  MoveL 4360 to (0, -14.4, 0.6) mm, rotated rx 0 ry 0 rz 180 deg; joints [18.174, -54.447, 108.401, -157.902, 56.008, 77.211]
  MoveL 4361 to (0, -15, 0.6) mm, rotated rx 0 ry 0 rz 180 deg; joints [18.174, -54.475, 108.395, -157.894, 55.977, 77.196]
  MoveL 4362 to (-200, -15, 0.6) mm, rotated rx 0 ry 0 rz 180 deg; joints [21.022, -63.449, 124.341, -156.258, 62.995, 78.705]
  MoveL 4363 to (-200, -15.6, 0.6) mm, rotated rx 0 ry 0 rz 180 deg; joints [21.022, -63.483, 124.335, -156.249, 62.958, 78.687]
  MoveL 4364 to (0, -15.6, 0.6) mm, rotated rx 0 ry 0 rz 180 deg; joints [18.174, -54.503, 108.39, -157.885, 55.945, 77.18]
  MoveL 4365 to (0, -16.2, 0.6) mm, rotated rx 0 ry 0 rz 180 deg; joints [18.174, -54.532, 108.384, -157.877, 55.914, 77.165]
  MoveL 4366 to (-200, -16.2, 0.6) mm, rotated rx 0 ry 0 rz 180 deg; joints [21.022, -63.518, 124.329, -156.241, 62.921, 78.669]
  MoveL 4367 to (-200, -16.8, 0.6) mm, rotated rx 0 ry 0 rz 180 deg; joints [21.022, -63.552, 124.323, -156.233, 62.883, 78.65]
  MoveL 4368 to (0, -16.8, 0.6) mm, rotated rx 0 ry 0 rz 180 deg; joints [18.174, -54.56, 108.378, -157.868, 55.882, 77.149]
  MoveL 4369 to (0, -17.4, 0.6) mm, rotated rx 0 ry 0 rz 180 deg; joints [18.174, -54.588, 108.373, -157.859, 55.851, 77.134]
  MoveL 4370 to (-200, -17.4, 0.6) mm, rotated rx 0 ry 0 rz 180 deg; joints [21.022, -63.586, 124.317, -156.224, 62.846, 78.632]
  MoveL 4371 to (-200, -18, 0.6) mm, rotated rx 0 ry 0 rz 180 deg; joints [21.022, -63.621, 124.311, -156.216, 62.809, 78.614]
  MoveL 4372 to (0, -18, 0.6) mm, rotated rx 0 ry 0 rz 180 deg; joints [18.174, -54.616, 108.367, -157.851, 55.819, 77.119]
  MoveL 4373 to (0, -18.6, 0.6) mm, rotated rx 0 ry 0 rz 180 deg; joints [18.174, -54.645, 108.361, -157.842, 55.788, 77.103]
  MoveL 4374 to (-200, -18.6, 0.6) mm, rotated rx 0 ry 0 rz 180 deg; joints [21.022, -63.655, 124.304, -156.208, 62.772, 78.595]
  MoveL 4375 to (-200, -19.2, 0.6) mm, rotated rx 0 ry 0 rz 180 deg; joints [21.022, -63.689, 124.298, -156.199, 62.735, 78.577]
  MoveL 4376 to (0, -19.2, 0.6) mm, rotated rx 0 ry 0 rz 180 deg; joints [18.174, -54.673, 108.355, -157.833, 55.756, 77.087]
  MoveL 4377 to (0, -19.8, 0.6) mm, rotated rx 0 ry 0 rz 180 deg; joints [18.174, -54.701, 108.349, -157.824, 55.725, 77.072]
  MoveL 4378 to (-200, -19.8, 0.6) mm, rotated rx 0 ry 0 rz 180 deg; joints [21.022, -63.724, 124.292, -156.191, 62.698, 78.558]
  MoveL 4379 to (-200, -20.4, 0.6) mm, rotated rx 0 ry 0 rz 180 deg; joints [21.022, -63.758, 124.285, -156.182, 62.661, 78.54]
  MoveL 4380 to (0, -20.4, 0.6) mm, rotated rx 0 ry 0 rz 180 deg; joints [18.174, -54.729, 108.344, -157.816, 55.693, 77.056]
  MoveL 4381 to (0, -21, 0.6) mm, rotated rx 0 ry 0 rz 180 deg; joints [18.174, -54.757, 108.338, -157.807, 55.662, 77.041]
  MoveL 4382 to (-200, -21, 0.6) mm, rotated rx 0 ry 0 rz 180 deg; joints [21.022, -63.792, 124.279, -156.174, 62.623, 78.521]
  MoveL 4383 to (-200, -21.6, 0.6) mm, rotated rx 0 ry 0 rz 180 deg; joints [21.022, -63.826, 124.272, -156.165, 62.586, 78.503]
  MoveL 4384 to (0, -21.6, 0.6) mm, rotated rx 0 ry 0 rz 180 deg; joints [18.174, -54.786, 108.332, -157.798, 55.63, 77.025]
  MoveL 4385 to (0, -22.2, 0.6) mm, rotated rx 0 ry 0 rz 180 deg; joints [18.174, -54.814, 108.326, -157.789, 55.599, 77.01]
  MoveL 4386 to (-200, -22.2, 0.6) mm, rotated rx 0 ry 0 rz 180 deg; joints [21.022, -63.86, 124.266, -156.157, 62.549, 78.484]
  MoveL 4387 to (-200, -22.8, 0.6) mm, rotated rx 0 ry 0 rz 180 deg; joints [21.022, -63.895, 124.26, -156.148, 62.512, 78.466]
  MoveL 4388 to (0, -22.8, 0.6) mm, rotated rx 0 ry 0 rz 180 deg; joints [18.174, -54.842, 108.32, -157.78, 55.567, 76.994]
  MoveL 4389 to (0, -23.4, 0.6) mm, rotated rx 0 ry 0 rz 180 deg; joints [18.174, -54.87, 108.314, -157.771, 55.535, 76.978]
  MoveL 4390 to (-200, -23.4, 0.6) mm, rotated rx 0 ry 0 rz 180 deg; joints [21.022, -63.929, 124.253, -156.14, 62.475, 78.447]
  MoveL 4391 to (-200, -24, 0.6) mm, rotated rx 0 ry 0 rz 180 deg; joints [21.022, -63.963, 124.246, -156.131, 62.438, 78.429]
  MoveL 4392 to (0, -24, 0.6) mm, rotated rx 0 ry 0 rz 180 deg; joints [18.174, -54.898, 108.308, -157.763, 55.504, 76.963]
  MoveL 4393 to (0, -24.6, 0.6) mm, rotated rx 0 ry 0 rz 180 deg; joints [18.174, -54.926, 108.302, -157.754, 55.472, 76.947]
  MoveL 4394 to (-200, -24.6, 0.6) mm, rotated rx 0 ry 0 rz 180 deg; joints [21.022, -63.997, 124.24, -156.122, 62.4, 78.41]
  MoveL 4395 to (-200, -25.2, 0.6) mm, rotated rx 0 ry 0 rz 180 deg; joints [21.022, -64.031, 124.233, -156.114, 62.363, 78.392]
  MoveL 4396 to (0, -25.2, 0.6) mm, rotated rx 0 ry 0 rz 180 deg; joints [18.174, -54.954, 108.296, -157.745, 55.441, 76.931]
  MoveL 4397 to (0, -25.8, 0.6) mm, rotated rx 0 ry 0 rz 180 deg; joints [18.174, -54.982, 108.289, -157.736, 55.409, 76.916]
  MoveL 4398 to (-200, -25.8, 0.6) mm, rotated rx 0 ry 0 rz 180 deg; joints [21.022, -64.065, 124.227, -156.105, 62.326, 78.373]
  MoveL 4399 to (-200, -26.4, 0.6) mm, rotated rx 0 ry 0 rz 180 deg; joints [21.022, -64.099, 124.22, -156.097, 62.289, 78.354]
  MoveL 4400 to (0, -26.4, 0.6) mm, rotated rx 0 ry 0 rz 180 deg; joints [18.174, -55.01, 108.283, -157.727, 55.377, 76.9]
  MoveL 4401 to (0, -27, 0.6) mm, rotated rx 0 ry 0 rz 180 deg; joints [18.174, -55.038, 108.277, -157.718, 55.346, 76.884]
  MoveL 4402 to (-200, -27, 0.6) mm, rotated rx 0 ry 0 rz 180 deg; joints [21.022, -64.133, 124.213, -156.088, 62.252, 78.336]
  MoveL 4403 to (-200, -27.6, 0.6) mm, rotated rx 0 ry 0 rz 180 deg; joints [21.022, -64.167, 124.206, -156.079, 62.214, 78.317]
  MoveL 4404 to (0, -27.6, 0.6) mm, rotated rx 0 ry 0 rz 180 deg; joints [18.174, -55.066, 108.271, -157.709, 55.314, 76.868]
  MoveL 4405 to (0, -28.2, 0.6) mm, rotated rx 0 ry 0 rz 180 deg; joints [18.174, -55.094, 108.265, -157.7, 55.282, 76.852]
  MoveL 4406 to (-200, -28.2, 0.6) mm, rotated rx 0 ry 0 rz 180 deg; joints [21.022, -64.201, 124.2, -156.07, 62.177, 78.298]
  MoveL 4407 to (-200, -28.8, 0.6) mm, rotated rx 0 ry 0 rz 180 deg; joints [21.022, -64.235, 124.193, -156.062, 62.14, 78.28]
  MoveL 4408 to (0, -28.8, 0.6) mm, rotated rx 0 ry 0 rz 180 deg; joints [18.174, -55.122, 108.258, -157.691, 55.251, 76.837]
  MoveL 4409 to (0, -29.4, 0.6) mm, rotated rx 0 ry 0 rz 180 deg; joints [18.174, -55.15, 108.252, -157.682, 55.219, 76.821]
  MoveL 4410 to (-200, -29.4, 0.6) mm, rotated rx 0 ry 0 rz 180 deg; joints [21.022, -64.269, 124.186, -156.053, 62.103, 78.261]
  MoveL 4411 to (-200, -30, 0.6) mm, rotated rx 0 ry 0 rz 180 deg; joints [21.022, -64.303, 124.179, -156.044, 62.065, 78.242]
  MoveL 4412 to (0, -30, 0.6) mm, rotated rx 0 ry 0 rz 180 deg; joints [18.174, -55.178, 108.246, -157.673, 55.187, 76.805]
  MoveL 4413 to (0, -30.6, 0.61) mm, rotated rx 2.39 ry 0 rz 180 deg; joints [18.094, -55.924, 108.131, -157.537, 54.374, 78.846]
  MoveL 4414 to (-200, -30.6, 0.61) mm, rotated rx 2.39 ry 0 rz 180 deg; joints [20.931, -65.205, 124.052, -155.918, 61.106, 80.201]
  MoveL 4415 to (-200, -31.2, 0.65) mm, rotated rx 4.78 ry 0 rz 180 deg; joints [20.813, -66.1, 123.923, -155.815, 60.147, 82.174]
  MoveL 4416 to (0, -31.2, 0.65) mm, rotated rx 4.78 ry 0 rz 180 deg; joints [17.989, -56.664, 108.016, -157.424, 53.559, 80.903]
  MoveL 4417 to (0, -31.8, 0.71) mm, rotated rx 7.16 ry 0 rz 180 deg; joints [17.861, -57.396, 107.901, -157.336, 52.745, 82.976]
  MoveL 4418 to (-200, -31.8, 0.71) mm, rotated rx 7.16 ry 0 rz 180 deg; joints [20.668, -66.984, 123.793, -155.736, 59.19, 84.161]
  MoveL 4419 to (-200, -32.39, 0.8) mm, rotated rx 9.55 ry 0 rz 180 deg; joints [20.495, -67.858, 123.663, -155.681, 58.234, 86.167]
  MoveL 4420 to (0, -32.39, 0.8) mm, rotated rx 9.55 ry 0 rz 180 deg; joints [17.708, -58.12, 107.785, -157.273, 51.933, 85.068]
  MoveL 4421 to (0, -32.98, 0.91) mm, rotated rx 11.94 ry 0 rz 180 deg; joints [17.531, -58.835, 107.67, -157.236, 51.122, 87.181]
  MoveL 4422 to (-200, -32.98, 0.91) mm, rotated rx 11.94 ry 0 rz 180 deg; joints [20.295, -68.721, 123.531, -155.653, 57.282, 88.193]
  MoveL 4423 to (-200, -33.56, 1.05) mm, rotated rx 14.32 ry 0 rz 180 deg; joints [20.068, -69.57, 123.4, -155.652, 56.333, 90.241]
  MoveL 4424 to (0, -33.56, 1.05) mm, rotated rx 14.32 ry 0 rz 180 deg; joints [17.331, -59.54, 107.555, -157.227, 50.315, 89.317]
  MoveL 4425 to (0, -34.14, 1.21) mm, rotated rx 16.71 ry 0 rz 180 deg; joints [17.107, -60.233, 107.441, -157.247, 49.513, 91.478]
  MoveL 4426 to (-200, -34.14, 1.21) mm, rotated rx 16.71 ry 0 rz 180 deg; joints [19.814, -70.405, 123.269, -155.68, 55.391, 92.314]
  MoveL 4427 to (-200, -34.71, 1.39) mm, rotated rx 19.1 ry 0 rz 180 deg; joints [19.533, -71.225, 123.138, -155.738, 54.454, 94.416]
  MoveL 4428 to (0, -34.71, 1.39) mm, rotated rx 19.1 ry 0 rz 180 deg; joints [16.859, -60.914, 107.328, -157.297, 48.715, 93.667]
  MoveL 4429 to (0, -35.27, 1.6) mm, rotated rx 21.49 ry 0 rz 180 deg; joints [16.589, -61.581, 107.218, -157.379, 47.925, 95.885]
  MoveL 4430 to (-200, -35.27, 1.6) mm, rotated rx 21.49 ry 0 rz 180 deg; joints [19.225, -72.028, 123.009, -155.827, 53.526, 96.546]
  MoveL 4431 to (-200, -35.83, 1.83) mm, rotated rx 23.87 ry 0 rz 180 deg; joints [18.892, -72.813, 122.882, -155.95, 52.606, 98.709]
  MoveL 4432 to (0, -35.83, 1.83) mm, rotated rx 23.87 ry 0 rz 180 deg; joints [16.295, -62.234, 107.109, -157.495, 47.142, 98.134]
  MoveL 4433 to (0, -36.37, 2.09) mm, rotated rx 26.26 ry 0 rz 180 deg; joints [15.979, -62.873, 107.003, -157.645, 46.368, 100.418]
  MoveL 4434 to (-200, -36.37, 2.09) mm, rotated rx 26.26 ry 0 rz 180 deg; joints [18.532, -73.58, 122.757, -156.107, 51.696, 100.907]
  MoveL 4435 to (-200, -36.9, 2.36) mm, rotated rx 28.65 ry 0 rz 180 deg; joints [18.147, -74.328, 122.635, -156.302, 50.798, 103.142]
  MoveL 4436 to (0, -36.9, 2.36) mm, rotated rx 28.65 ry 0 rz 180 deg; joints [15.641, -63.494, 106.9, -157.832, 45.604, 102.738]
  MoveL 4437 to (0, -37.42, 2.66) mm, rotated rx 31.03 ry 0 rz 180 deg; joints [15.281, -64.099, 106.8, -158.057, 44.853, 105.095]
  MoveL 4438 to (-200, -37.42, 2.66) mm, rotated rx 31.03 ry 0 rz 180 deg; joints [17.737, -75.054, 122.516, -156.535, 49.913, 105.418]
  MoveL 4439 to (-200, -37.93, 2.98) mm, rotated rx 33.42 ry 0 rz 180 deg; joints [17.301, -75.76, 122.401, -156.809, 49.042, 107.737]
  MoveL 4440 to (0, -37.93, 2.98) mm, rotated rx 33.42 ry 0 rz 180 deg; joints [14.9, -64.687, 106.705, -158.321, 44.114, 107.494]
  MoveL 4441 to (0, -38.42, 3.32) mm, rotated rx 35.81 ry 0 rz 180 deg; joints [14.498, -65.256, 106.613, -158.627, 43.39, 109.935]
  MoveL 4442 to (-200, -38.42, 3.32) mm, rotated rx 35.81 ry 0 rz 180 deg; joints [16.842, -76.442, 122.29, -157.125, 48.188, 110.1]
  MoveL 4443 to (-200, -38.91, 3.68) mm, rotated rx 38.2 ry 0 rz 180 deg; joints [16.358, -77.102, 122.185, -157.486, 47.352, 112.511]
  MoveL 4444 to (0, -38.91, 3.68) mm, rotated rx 38.2 ry 0 rz 180 deg; joints [14.076, -65.805, 106.527, -158.976, 42.682, 112.42]
  MoveL 4445 to (0, -39.37, 4.06) mm, rotated rx 40.59 ry 0 rz 180 deg; joints [13.634, -66.334, 106.446, -159.37, 41.992, 114.953]
  MoveL 4446 to (-200, -39.37, 4.06) mm, rotated rx 40.59 ry 0 rz 180 deg; joints [15.852, -77.737, 122.085, -157.893, 46.535, 114.973]
  MoveL 4447 to (-200, -39.82, 4.46) mm, rotated rx 42.97 ry 0 rz 180 deg; joints [15.322, -78.347, 121.991, -158.348, 45.739, 117.486]
  MoveL 4448 to (0, -39.82, 4.46) mm, rotated rx 42.97 ry 0 rz 180 deg; joints [13.173, -66.843, 106.37, -159.81, 41.321, 117.533]
  MoveL 4449 to (0, -40.25, 4.88) mm, rotated rx 45.36 ry 0 rz 180 deg; joints [12.693, -67.329, 106.301, -160.297, 40.672, 120.163]
  MoveL 4450 to (-200, -40.25, 4.88) mm, rotated rx 45.36 ry 0 rz 180 deg; joints [14.771, -78.931, 121.903, -158.853, 44.968, 120.054]
  MoveL 4451 to (-200, -40.66, 5.32) mm, rotated rx 47.75 ry 0 rz 180 deg; joints [14.199, -79.488, 121.823, -159.409, 44.222, 122.677]
  MoveL 4452 to (0, -40.66, 5.32) mm, rotated rx 47.75 ry 0 rz 180 deg; joints [12.196, -67.794, 106.238, -160.832, 40.045, 122.844]
  MoveL 4453 to (0, -41.05, 5.77) mm, rotated rx 50.13 ry 0 rz 180 deg; joints [11.681, -68.236, 106.182, -161.417, 39.444, 125.579]
  MoveL 4454 to (-200, -41.05, 5.77) mm, rotated rx 50.13 ry 0 rz 180 deg; joints [13.605, -80.018, 121.75, -160.019, 43.504, 125.36]
  MoveL 4455 to (-200, -41.43, 6.24) mm, rotated rx 52.52 ry 0 rz 180 deg; joints [12.993, -80.519, 121.685, -160.682, 42.817, 128.101]
  MoveL 4456 to (0, -41.43, 6.24) mm, rotated rx 52.52 ry 0 rz 180 deg; joints [11.15, -68.654, 106.134, -162.052, 38.869, 128.366]
  MoveL 4457 to (0, -41.78, 6.72) mm, rotated rx 54.91 ry 0 rz 180 deg; joints [10.604, -69.047, 106.093, -162.737, 38.324, 131.207]
  MoveL 4458 to (-200, -41.78, 6.72) mm, rotated rx 54.91 ry 0 rz 180 deg; joints [12.362, -80.992, 121.629, -161.4, 42.162, 130.901]
  MoveL 4459 to (-200, -42.12, 7.22) mm, rotated rx 57.3 ry 0 rz 180 deg; joints [11.713, -81.435, 121.582, -162.174, 41.541, 133.763]
  MoveL 4460 to (0, -42.12, 7.22) mm, rotated rx 57.3 ry 0 rz 180 deg; joints [10.043, -69.416, 106.061, -163.472, 37.809, 134.102]
  MoveL 4461 to (0, -42.43, 7.73) mm, rotated rx 59.68 ry 0 rz 180 deg; joints [9.469, -69.76, 106.037, -164.257, 37.327, 137.048]
  MoveL 4462 to (-200, -42.43, 7.73) mm, rotated rx 59.68 ry 0 rz 180 deg; joints [11.048, -81.848, 121.544, -163.002, 40.959, 136.684]
  MoveL 4463 to (-200, -42.72, 8.26) mm, rotated rx 62.07 ry 0 rz 180 deg; joints [10.368, -82.229, 121.516, -163.884, 40.416, 139.663]
  MoveL 4464 to (0, -42.72, 8.26) mm, rotated rx 62.07 ry 0 rz 180 deg; joints [8.883, -70.078, 106.021, -165.091, 36.88, 140.047]
  MoveL 4465 to (0, -42.99, 8.79) mm, rotated rx 64.46 ry 0 rz 180 deg; joints [8.284, -70.37, 106.015, -165.972, 36.47, 143.097]
  MoveL 4466 to (-200, -42.99, 8.79) mm, rotated rx 64.46 ry 0 rz 180 deg; joints [9.673, -82.58, 121.498, -164.82, 39.916, 142.702]
  MoveL 4467 to (-200, -43.24, 9.34) mm, rotated rx 66.84 ry 0 rz 180 deg; joints [8.965, -82.898, 121.49, -165.806, 39.461, 145.796]
  MoveL 4468 to (0, -43.24, 9.34) mm, rotated rx 66.84 ry 0 rz 180 deg; joints [7.675, -70.634, 106.017, -166.898, 36.099, 146.195]
  MoveL 4469 to (0, -43.46, 9.89) mm, rotated rx 69.23 ry 0 rz 180 deg; joints [7.057, -70.872, 106.029, -167.866, 35.769, 149.337]
  MoveL 4470 to (-200, -43.46, 9.89) mm, rotated rx 69.23 ry 0 rz 180 deg; joints [8.246, -83.184, 121.493, -166.841, 39.053, 148.942]
  MoveL 4471 to (-200, -43.66, 10.46) mm, rotated rx 71.62 ry 0 rz 180 deg; joints [7.517, -83.436, 121.507, -167.922, 38.695, 152.139]
  MoveL 4472 to (0, -43.66, 10.46) mm, rotated rx 71.62 ry 0 rz 180 deg; joints [6.431, -71.082, 106.051, -168.874, 35.481, 152.522]
  MoveL 4473 to (0, -43.84, 11.03) mm, rotated rx 74.01 ry 0 rz 180 deg; joints [5.797, -71.264, 106.082, -169.917, 35.237, 155.743]
  MoveL 4474 to (-200, -43.84, 11.03) mm, rotated rx 74.01 ry 0 rz 180 deg; joints [6.778, -83.656, 121.532, -169.044, 38.388, 155.379]
  MoveL 4475 to (-200, -44, 11.61) mm, rotated rx 76.39 ry 0 rz 180 deg; joints [6.032, -83.841, 121.568, -170.201, 38.135, 158.658]
  MoveL 4476 to (0, -44, 11.61) mm, rotated rx 76.39 ry 0 rz 180 deg; joints [5.158, -71.418, 106.123, -170.991, 35.039, 158.997]
  MoveL 4477 to (0, -44.12, 12.2) mm, rotated rx 78.78 ry 0 rz 180 deg; joints [4.514, -71.543, 106.173, -172.09, 34.887, 162.28]
  MoveL 4478 to (-200, -44.12, 12.2) mm, rotated rx 78.78 ry 0 rz 180 deg; joints [5.281, -83.992, 121.615, -171.391, 37.938, 161.973]
  MoveL 4479 to (-200, -44.23, 12.79) mm, rotated rx 81.17 ry 0 rz 180 deg; joints [4.525, -84.109, 121.674, -172.604, 37.797, 165.313]
  MoveL 4480 to (0, -44.23, 12.79) mm, rotated rx 81.17 ry 0 rz 180 deg; joints [3.867, -71.639, 106.234, -173.21, 34.783, 165.584]
  MoveL 4481 to (0, -44.31, 13.38) mm, rotated rx 83.56 ry 0 rz 180 deg; joints [3.218, -71.706, 106.304, -174.345, 34.728, 168.903]
  MoveL 4482 to (-200, -44.31, 13.38) mm, rotated rx 83.56 ry 0 rz 180 deg; joints [3.766, -84.191, 121.744, -173.836, 37.714, 168.673]
  MoveL 4483 to (-200, -44.36, 13.98) mm, rotated rx 85.94 ry 0 rz 180 deg; joints [3.006, -84.237, 121.825, -175.08, 37.69, 172.047]
  MoveL 4484 to (0, -44.36, 13.98) mm, rotated rx 85.94 ry 0 rz 180 deg; joints [2.568, -71.744, 106.384, -175.488, 34.722, 172.233]
  MoveL 4485 to (0, -44.39, 14.58) mm, rotated rx 88.33 ry 0 rz 180 deg; joints [1.919, -71.753, 106.473, -176.633, 34.766, 175.564]
  MoveL 4486 to (-200, -44.39, 14.58) mm, rotated rx 88.33 ry 0 rz 180 deg; joints [2.246, -84.249, 121.918, -176.328, 37.726, 175.425]
  MoveL 4487 to (-200, -44.4, 15.18) mm, rotated rx 90 ry 0 rz 180 deg; joints [1.707, -84.236, 121.989, -177.213, 37.786, 177.797]
  MoveL 4488 to (0, -44.4, 15.18) mm, rotated rx 90 ry 0 rz 180 deg; joints [1.459, -71.742, 106.541, -177.445, 34.826, 177.903]
  MoveL 4489 to (0, -44.4, 15.78) mm, rotated rx 90 ry 0 rz 180 deg; joints [1.433, -71.743, 106.542, -177.489, 34.825, 177.939]
  MoveL 4490 to (-200, -44.4, 15.78) mm, rotated rx 90 ry 0 rz 180 deg; joints [1.678, -84.237, 121.99, -177.261, 37.785, 177.834]
  MoveL 4491 to (-200, -44.4, 16.38) mm, rotated rx 90 ry 0 rz 180 deg; joints [1.649, -84.239, 121.992, -177.308, 37.784, 177.872]
  MoveL 4492 to (0, -44.4, 16.38) mm, rotated rx 90 ry 0 rz 180 deg; joints [1.408, -71.744, 106.544, -177.533, 34.825, 177.975]
  MoveL 4493 to (0, -44.4, 16.98) mm, rotated rx 90 ry 0 rz 180 deg; joints [1.383, -71.745, 106.545, -177.577, 34.824, 178.011]
  MoveL 4494 to (-200, -44.4, 16.98) mm, rotated rx 90 ry 0 rz 180 deg; joints [1.619, -84.24, 121.993, -177.356, 37.783, 177.91]
  MoveL 4495 to (-200, -44.4, 17.58) mm, rotated rx 90 ry 0 rz 180 deg; joints [1.59, -84.241, 121.994, -177.404, 37.782, 177.948]
  MoveL 4496 to (0, -44.4, 17.58) mm, rotated rx 90 ry 0 rz 180 deg; joints [1.358, -71.746, 106.546, -177.621, 34.824, 178.047]
  MoveL 4497 to (0, -44.4, 18.18) mm, rotated rx 90 ry 0 rz 180 deg; joints [1.333, -71.746, 106.547, -177.665, 34.823, 178.083]
  MoveL 4498 to (-200, -44.4, 18.18) mm, rotated rx 90 ry 0 rz 180 deg; joints [1.561, -84.242, 121.995, -177.452, 37.781, 177.986]
  MoveL 4499 to (-200, -44.4, 18.78) mm, rotated rx 90 ry 0 rz 180 deg; joints [1.531, -84.243, 121.996, -177.5, 37.78, 178.023]
  MoveL 4500 to (0, -44.4, 18.78) mm, rotated rx 90 ry 0 rz 180 deg; joints [1.308, -71.747, 106.548, -177.709, 34.823, 178.119]
  MoveL 4501 to (0, -44.4, 19.38) mm, rotated rx 90 ry 0 rz 180 deg; joints [1.283, -71.748, 106.549, -177.752, 34.822, 178.155]
  MoveL 4502 to (-200, -44.4, 19.38) mm, rotated rx 90 ry 0 rz 180 deg; joints [1.502, -84.244, 121.998, -177.548, 37.779, 178.061]
  MoveL 4503 to (-200, -44.4, 19.98) mm, rotated rx 90 ry 0 rz 180 deg; joints [1.473, -84.245, 121.999, -177.595, 37.778, 178.099]
  MoveL 4504 to (0, -44.4, 19.98) mm, rotated rx 90 ry 0 rz 180 deg; joints [1.258, -71.749, 106.551, -177.796, 34.822, 178.191]
  MoveL 4505 to (0, -44.4, 20.58) mm, rotated rx 90 ry 0 rz 180 deg; joints [1.233, -71.75, 106.552, -177.84, 34.821, 178.227]
  MoveL 4506 to (-200, -44.4, 20.58) mm, rotated rx 90 ry 0 rz 180 deg; joints [1.443, -84.246, 122, -177.643, 37.777, 178.137]
  MoveL 4507 to (-200, -44.4, 21.18) mm, rotated rx 90 ry 0 rz 180 deg; joints [1.414, -84.247, 122.001, -177.691, 37.777, 178.175]
  MoveL 4508 to (0, -44.4, 21.18) mm, rotated rx 90 ry 0 rz 180 deg; joints [1.208, -71.75, 106.553, -177.884, 34.821, 178.263]
  MoveL 4509 to (0, -44.4, 21.78) mm, rotated rx 90 ry 0 rz 180 deg; joints [1.183, -71.751, 106.554, -177.928, 34.82, 178.299]
  MoveL 4510 to (-200, -44.4, 21.78) mm, rotated rx 90 ry 0 rz 180 deg; joints [1.385, -84.248, 122.002, -177.739, 37.776, 178.212]
  MoveL 4511 to (-200, -44.4, 22.38) mm, rotated rx 90 ry 0 rz 180 deg; joints [1.356, -84.249, 122.003, -177.787, 37.775, 178.25]
  MoveL 4512 to (0, -44.4, 22.38) mm, rotated rx 90 ry 0 rz 180 deg; joints [1.158, -71.752, 106.555, -177.972, 34.82, 178.335]
  MoveL 4513 to (0, -44.4, 22.98) mm, rotated rx 90 ry 0 rz 180 deg; joints [1.133, -71.753, 106.556, -178.016, 34.819, 178.371]
  MoveL 4514 to (-200, -44.4, 22.98) mm, rotated rx 90 ry 0 rz 180 deg; joints [1.326, -84.25, 122.004, -177.835, 37.774, 178.288]
  MoveL 4515 to (-200, -44.4, 23.58) mm, rotated rx 90 ry 0 rz 180 deg; joints [1.297, -84.25, 122.005, -177.882, 37.773, 178.326]
  MoveL 4516 to (0, -44.4, 23.58) mm, rotated rx 90 ry 0 rz 180 deg; joints [1.108, -71.753, 106.557, -178.059, 34.819, 178.407]
  MoveL 4517 to (0, -44.4, 24.18) mm, rotated rx 90 ry 0 rz 180 deg; joints [1.083, -71.754, 106.558, -178.103, 34.818, 178.443]
  MoveL 4518 to (-200, -44.4, 24.18) mm, rotated rx 90 ry 0 rz 180 deg; joints [1.268, -84.251, 122.006, -177.93, 37.773, 178.364]
  MoveL 4519 to (-200, -44.4, 24.78) mm, rotated rx 90 ry 0 rz 180 deg; joints [1.238, -84.252, 122.007, -177.978, 37.772, 178.402]
  MoveL 4520 to (0, -44.4, 24.78) mm, rotated rx 90 ry 0 rz 180 deg; joints [1.058, -71.755, 106.559, -178.147, 34.818, 178.479]
  MoveL 4521 to (0, -44.4, 25.38) mm, rotated rx 90 ry 0 rz 180 deg; joints [1.033, -71.756, 106.56, -178.191, 34.817, 178.515]
  MoveL 4522 to (-200, -44.4, 25.38) mm, rotated rx 90 ry 0 rz 180 deg; joints [1.209, -84.253, 122.008, -178.026, 37.771, 178.439]
  MoveL 4523 to (-200, -44.4, 25.98) mm, rotated rx 90 ry 0 rz 180 deg; joints [1.18, -84.254, 122.009, -178.074, 37.77, 178.477]
  MoveL 4524 to (0, -44.4, 25.98) mm, rotated rx 90 ry 0 rz 180 deg; joints [1.008, -71.756, 106.56, -178.235, 34.817, 178.551]
  MoveL 4525 to (0, -44.4, 26.58) mm, rotated rx 90 ry 0 rz 180 deg; joints [0.983, -71.757, 106.561, -178.279, 34.817, 178.587]
  MoveL 4526 to (-200, -44.4, 26.58) mm, rotated rx 90 ry 0 rz 180 deg; joints [1.15, -84.255, 122.009, -178.122, 37.77, 178.515]
  MoveL 4527 to (-200, -44.4, 27.18) mm, rotated rx 90 ry 0 rz 180 deg; joints [1.121, -84.255, 122.01, -178.17, 37.769, 178.553]
  MoveL 4528 to (0, -44.4, 27.18) mm, rotated rx 90 ry 0 rz 180 deg; joints [0.958, -71.757, 106.562, -178.323, 34.816, 178.623]
  MoveL 4529 to (0, -44.4, 27.78) mm, rotated rx 90 ry 0 rz 180 deg; joints [0.933, -71.758, 106.563, -178.366, 34.816, 178.659]
  MoveL 4530 to (-200, -44.4, 27.78) mm, rotated rx 90 ry 0 rz 180 deg; joints [1.092, -84.256, 122.011, -178.217, 37.768, 178.591]
  MoveL 4531 to (-200, -44.4, 28.38) mm, rotated rx 90 ry 0 rz 180 deg; joints [1.062, -84.257, 122.012, -178.265, 37.768, 178.629]
  MoveL 4532 to (0, -44.4, 28.38) mm, rotated rx 90 ry 0 rz 180 deg; joints [0.907, -71.759, 106.564, -178.41, 34.815, 178.695]
  MoveL 4533 to (0, -44.4, 28.98) mm, rotated rx 90 ry 0 rz 180 deg; joints [0.882, -71.759, 106.565, -178.454, 34.815, 178.731]
  MoveL 4534 to (-200, -44.4, 28.98) mm, rotated rx 90 ry 0 rz 180 deg; joints [1.033, -84.258, 122.013, -178.313, 37.767, 178.666]
  MoveL 4535 to (-200, -44.4, 29.58) mm, rotated rx 90 ry 0 rz 180 deg; joints [1.004, -84.258, 122.014, -178.361, 37.767, 178.704]
  MoveL 4536 to (0, -44.4, 29.58) mm, rotated rx 90 ry 0 rz 180 deg; joints [0.857, -71.76, 106.565, -178.498, 34.815, 178.767]
  MoveL 4537 to (0, -44.4, 30.18) mm, rotated rx 90 ry 0 rz 180 deg; joints [0.832, -71.76, 106.566, -178.542, 34.814, 178.803]
  MoveL 4538 to (-200, -44.4, 30.18) mm, rotated rx 90 ry 0 rz 180 deg; joints [0.974, -84.259, 122.014, -178.409, 37.766, 178.742]
  MoveL 4539 to (-200, -44.4, 30.78) mm, rotated rx 90 ry 0 rz 180 deg; joints [0.945, -84.26, 122.015, -178.457, 37.766, 178.78]
  MoveL 4540 to (0, -44.4, 30.78) mm, rotated rx 90 ry 0 rz 180 deg; joints [0.807, -71.761, 106.567, -178.586, 34.814, 178.839]
  MoveL 4541 to (0, -44.4, 31.38) mm, rotated rx 90 ry 0 rz 180 deg; joints [0.782, -71.761, 106.567, -178.63, 34.814, 178.875]
  MoveL 4542 to (-200, -44.4, 31.38) mm, rotated rx 90 ry 0 rz 180 deg; joints [0.916, -84.26, 122.016, -178.505, 37.765, 178.818]
  MoveL 4543 to (-200, -44.4, 31.98) mm, rotated rx 90 ry 0 rz 180 deg; joints [0.886, -84.261, 122.016, -178.553, 37.764, 178.856]
  MoveL 4544 to (0, -44.4, 31.98) mm, rotated rx 90 ry 0 rz 180 deg; joints [0.757, -71.762, 106.568, -178.674, 34.813, 178.911]
  MoveL 4545 to (0, -44.4, 32.58) mm, rotated rx 90 ry 0 rz 180 deg; joints [0.732, -71.762, 106.569, -178.718, 34.813, 178.947]
  MoveL 4546 to (-200, -44.4, 32.58) mm, rotated rx 90 ry 0 rz 180 deg; joints [0.857, -84.261, 122.017, -178.6, 37.764, 178.894]
  MoveL 4547 to (-200, -44.4, 33.18) mm, rotated rx 90 ry 0 rz 180 deg; joints [0.828, -84.262, 122.018, -178.648, 37.763, 178.931]
  MoveL 4548 to (0, -44.4, 33.18) mm, rotated rx 90 ry 0 rz 180 deg; joints [0.707, -71.763, 106.569, -178.761, 34.813, 178.983]
  MoveL 4549 to (0, -44.4, 33.78) mm, rotated rx 90 ry 0 rz 180 deg; joints [0.682, -71.763, 106.57, -178.805, 34.813, 179.019]
  MoveL 4550 to (-200, -44.4, 33.78) mm, rotated rx 90 ry 0 rz 180 deg; joints [0.798, -84.262, 122.018, -178.696, 37.763, 178.969]
  MoveL 4551 to (-200, -44.4, 34.38) mm, rotated rx 90 ry 0 rz 180 deg; joints [0.769, -84.263, 122.019, -178.744, 37.763, 179.007]
  MoveL 4552 to (0, -44.4, 34.38) mm, rotated rx 90 ry 0 rz 180 deg; joints [0.657, -71.764, 106.571, -178.849, 34.812, 179.055]
  MoveL 4553 to (0, -44.4, 34.98) mm, rotated rx 90 ry 0 rz 180 deg; joints [0.632, -71.764, 106.571, -178.893, 34.812, 179.091]
  MoveL 4554 to (-200, -44.4, 34.98) mm, rotated rx 90 ry 0 rz 180 deg; joints [0.74, -84.263, 122.019, -178.792, 37.762, 179.045]
  MoveL 4555 to (-200, -44.4, 35.58) mm, rotated rx 90 ry 0 rz 180 deg; joints [0.71, -84.264, 122.02, -178.84, 37.762, 179.083]
  MoveL 4556 to (0, -44.4, 35.58) mm, rotated rx 90 ry 0 rz 180 deg; joints [0.607, -71.765, 106.572, -178.937, 34.812, 179.127]
  MoveL 4557 to (0, -44.4, 36.18) mm, rotated rx 90 ry 0 rz 180 deg; joints [0.582, -71.765, 106.572, -178.981, 34.812, 179.163]
  MoveL 4558 to (-200, -44.4, 36.18) mm, rotated rx 90 ry 0 rz 180 deg; joints [0.681, -84.264, 122.02, -178.888, 37.761, 179.121]
  MoveL 4559 to (-200, -44.4, 36.78) mm, rotated rx 90 ry 0 rz 180 deg; joints [0.652, -84.265, 122.021, -178.936, 37.761, 179.159]
  MoveL 4560 to (0, -44.4, 36.78) mm, rotated rx 90 ry 0 rz 180 deg; joints [0.557, -71.765, 106.573, -179.025, 34.811, 179.199]
  MoveL 4561 to (0, -44.4, 37.38) mm, rotated rx 90 ry 0 rz 180 deg; joints [0.532, -71.766, 106.573, -179.069, 34.811, 179.235]
  MoveL 4562 to (-200, -44.4, 37.38) mm, rotated rx 90 ry 0 rz 180 deg; joints [0.622, -84.265, 122.021, -178.984, 37.76, 179.196]
  MoveL 4563 to (-200, -44.4, 37.98) mm, rotated rx 90 ry 0 rz 180 deg; joints [0.593, -84.266, 122.022, -179.031, 37.76, 179.234]
  MoveL 4564 to (0, -44.4, 37.98) mm, rotated rx 90 ry 0 rz 180 deg; joints [0.507, -71.766, 106.574, -179.112, 34.811, 179.271]
  MoveL 4565 to (0, -44.4, 38.58) mm, rotated rx 90 ry 0 rz 180 deg; joints [0.482, -71.766, 106.574, -179.156, 34.811, 179.307]
  MoveL 4566 to (-200, -44.4, 38.58) mm, rotated rx 90 ry 0 rz 180 deg; joints [0.564, -84.266, 122.022, -179.079, 37.76, 179.272]
  MoveL 4567 to (-200, -44.4, 39.18) mm, rotated rx 90 ry 0 rz 180 deg; joints [0.534, -84.266, 122.023, -179.127, 37.759, 179.31]
  MoveL 4568 to (0, -44.4, 39.18) mm, rotated rx 90 ry 0 rz 180 deg; joints [0.457, -71.767, 106.574, -179.2, 34.81, 179.343]
  MoveL 4569 to (0, -44.4, 39.78) mm, rotated rx 90 ry 0 rz 180 deg; joints [0.431, -71.767, 106.575, -179.244, 34.81, 179.379]
  MoveL 4570 to (-200, -44.4, 39.78) mm, rotated rx 90 ry 0 rz 180 deg; joints [0.505, -84.267, 122.023, -179.175, 37.759, 179.348]
  MoveL 4571 to (-200, -44.4, 40.38) mm, rotated rx 90 ry 0 rz 180 deg; joints [0.476, -84.267, 122.024, -179.223, 37.759, 179.386]
  MoveL 4572 to (0, -44.4, 40.38) mm, rotated rx 90 ry 0 rz 180 deg; joints [0.406, -71.767, 106.575, -179.288, 34.81, 179.415]
  MoveL 4573 to (0, -44.4, 40.98) mm, rotated rx 90 ry 0 rz 180 deg; joints [0.381, -71.767, 106.576, -179.332, 34.81, 179.451]
  MoveL 4574 to (-200, -44.4, 40.98) mm, rotated rx 90 ry 0 rz 180 deg; joints [0.446, -84.267, 122.024, -179.271, 37.759, 179.424]
  MoveL 4575 to (-200, -44.4, 41.58) mm, rotated rx 90 ry 0 rz 180 deg; joints [0.417, -84.268, 122.024, -179.319, 37.758, 179.461]
  MoveL 4576 to (0, -44.4, 41.58) mm, rotated rx 90 ry 0 rz 180 deg; joints [0.356, -71.768, 106.576, -179.376, 34.81, 179.488]
  MoveL 4577 to (0, -44.4, 42.18) mm, rotated rx 90 ry 0 rz 180 deg; joints [0.331, -71.768, 106.576, -179.42, 34.81, 179.524]
  MoveL 4578 to (-200, -44.4, 42.18) mm, rotated rx 90 ry 0 rz 180 deg; joints [0.388, -84.268, 122.024, -179.367, 37.758, 179.499]
  MoveL 4579 to (-200, -44.4, 42.78) mm, rotated rx 90 ry 0 rz 180 deg; joints [0.358, -84.268, 122.025, -179.415, 37.758, 179.537]
  MoveL 4580 to (0, -44.4, 42.78) mm, rotated rx 90 ry 0 rz 180 deg; joints [0.306, -71.768, 106.576, -179.464, 34.81, 179.56]
  MoveL 4581 to (0, -44.4, 43.38) mm, rotated rx 90 ry 0 rz 180 deg; joints [0.281, -71.768, 106.577, -179.508, 34.809, 179.596]
  MoveL 4582 to (-200, -44.4, 43.38) mm, rotated rx 90 ry 0 rz 180 deg; joints [0.329, -84.269, 122.025, -179.463, 37.758, 179.575]
  MoveL 4583 to (-200, -44.4, 43.98) mm, rotated rx 90 ry 0 rz 180 deg; joints [0.3, -84.269, 122.025, -179.51, 37.758, 179.613]
  MoveL 4584 to (0, -44.4, 43.98) mm, rotated rx 90 ry 0 rz 180 deg; joints [0.256, -71.768, 106.577, -179.551, 34.809, 179.632]
  MoveL 4585 to (0, -44.4, 44.58) mm, rotated rx 90 ry 0 rz 180 deg; joints [0.231, -71.769, 106.577, -179.595, 34.809, 179.668]
  MoveL 4586 to (-200, -44.4, 44.58) mm, rotated rx 90 ry 0 rz 180 deg; joints [0.27, -84.269, 122.025, -179.558, 37.757, 179.651]
  MoveL 4587 to (-200, -44.4, 45.18) mm, rotated rx 90.72 ry 0 rz 180 deg; joints [0.022, -84.25, 122.049, -179.964, 37.799, -179.311]
  MoveL 4588 to (0, -44.4, 45.18) mm, rotated rx 90.72 ry 0 rz 180 deg; joints [0.019, -71.753, 106.599, -179.967, 34.846, -179.309]
  MoveL 4589 to (0, -44.38, 45.78) mm, rotated rx 93.11 ry 0 rz 180 deg; joints [-0.626, -71.682, 106.679, 178.909, 35.002, -176]
  MoveL 4590 to (-200, -44.38, 45.78) mm, rotated rx 93.11 ry 0 rz 180 deg; joints [-0.732, -84.166, 122.135, 178.81, 37.975, -175.956]
  MoveL 4591 to (-200, -44.33, 46.38) mm, rotated rx 95.49 ry 0 rz 180 deg; joints [-1.481, -84.045, 122.231, 177.605, 38.21, -172.625]
  MoveL 4592 to (0, -44.33, 46.38) mm, rotated rx 95.49 ry 0 rz 180 deg; joints [-1.265, -71.581, 106.767, 177.805, 35.206, -172.713]
  MoveL 4593 to (0, -44.26, 46.97) mm, rotated rx 97.88 ry 0 rz 180 deg; joints [-1.899, -71.451, 106.864, 176.725, 35.457, -169.452]
  MoveL 4594 to (-200, -44.26, 46.97) mm, rotated rx 97.88 ry 0 rz 180 deg; joints [-2.223, -83.89, 122.337, 176.428, 38.502, -169.323]
  MoveL 4595 to (-200, -44.17, 47.57) mm, rotated rx 100.27 ry 0 rz 180 deg; joints [-2.956, -83.699, 122.453, 175.284, 38.849, -166.056]
  MoveL 4596 to (0, -44.17, 47.57) mm, rotated rx 100.27 ry 0 rz 180 deg; joints [-2.526, -71.292, 106.97, 175.675, 35.755, -166.22]
  MoveL 4597 to (0, -44.05, 48.16) mm, rotated rx 102.66 ry 0 rz 180 deg; joints [-3.144, -71.104, 107.083, 174.659, 36.097, -163.025]
  MoveL 4598 to (-200, -44.05, 48.16) mm, rotated rx 102.66 ry 0 rz 180 deg; joints [-3.679, -83.474, 122.579, 174.18, 39.251, -162.832]
  MoveL 4599 to (-200, -43.91, 48.74) mm, rotated rx 105.04 ry 0 rz 180 deg; joints [-4.39, -83.213, 122.714, 173.119, 39.704, -159.653]
  MoveL 4600 to (0, -43.91, 48.74) mm, rotated rx 105.04 ry 0 rz 180 deg; joints [-3.752, -70.887, 107.204, 173.682, 36.483, -159.871]
  MoveL 4601 to (0, -43.74, 49.31) mm, rotated rx 107.43 ry 0 rz 180 deg; joints [-4.349, -70.642, 107.333, 172.745, 36.912, -156.758]
  MoveL 4602 to (-200, -43.74, 49.31) mm, rotated rx 107.43 ry 0 rz 180 deg; joints [-5.088, -82.918, 122.857, 172.104, 40.208, -156.524]
  MoveL 4603 to (-200, -43.55, 49.88) mm, rotated rx 109.82 ry 0 rz 180 deg; joints [-5.772, -82.589, 123.009, 171.139, 40.76, -153.448]
  MoveL 4604 to (0, -43.55, 49.88) mm, rotated rx 109.82 ry 0 rz 180 deg; joints [-4.935, -70.368, 107.468, 171.854, 37.379, -153.694]
  MoveL 4605 to (0, -43.33, 50.44) mm, rotated rx 112.2 ry 0 rz 180 deg; joints [-5.508, -70.067, 107.609, 171.008, 37.885, -150.677]
  MoveL 4606 to (-200, -43.33, 50.44) mm, rotated rx 112.2 ry 0 rz 180 deg; joints [-6.44, -82.226, 123.168, 170.227, 41.357, -150.429]
  MoveL 4607 to (-200, -43.09, 50.99) mm, rotated rx 114.59 ry 0 rz 180 deg; joints [-7.092, -81.829, 123.334, 169.367, 41.997, -147.465]
  MoveL 4608 to (0, -43.09, 50.99) mm, rotated rx 114.59 ry 0 rz 180 deg; joints [-6.066, -69.737, 107.756, 170.21, 38.428, -147.71]
  MoveL 4609 to (0, -42.83, 51.53) mm, rotated rx 116.98 ry 0 rz 180 deg; joints [-6.61, -69.381, 107.909, 169.462, 39.004, -144.795]
  MoveL 4610 to (-200, -42.83, 51.53) mm, rotated rx 116.98 ry 0 rz 180 deg; joints [-7.725, -81.4, 123.506, 168.563, 42.678, -144.561]
  MoveL 4611 to (-200, -42.55, 52.06) mm, rotated rx 119.37 ry 0 rz 180 deg; joints [-8.339, -80.938, 123.684, 167.814, 43.397, -141.716]
  MoveL 4612 to (0, -42.55, 52.06) mm, rotated rx 119.37 ry 0 rz 180 deg; joints [-7.137, -68.998, 108.066, 168.763, 39.612, -141.932]
  MoveL 4613 to (0, -42.24, 52.58) mm, rotated rx 121.75 ry 0 rz 180 deg; joints [-7.648, -68.588, 108.228, 168.114, 40.251, -139.12]
  MoveL 4614 to (-200, -42.24, 52.58) mm, rotated rx 121.75 ry 0 rz 180 deg; joints [-8.933, -80.444, 123.867, 167.119, 44.152, -138.928]
  MoveL 4615 to (-200, -41.92, 53.08) mm, rotated rx 124.14 ry 0 rz 180 deg; joints [-9.506, -79.918, 124.054, 166.479, 44.941, -136.199]
  MoveL 4616 to (0, -41.92, 53.08) mm, rotated rx 124.14 ry 0 rz 180 deg; joints [-8.141, -68.153, 108.393, 167.514, 40.917, -136.36]
  MoveL 4617 to (0, -41.57, 53.57) mm, rotated rx 126.53 ry 0 rz 180 deg; joints [-8.615, -67.692, 108.561, 166.963, 41.61, -133.65]
  MoveL 4618 to (-200, -41.57, 53.57) mm, rotated rx 126.53 ry 0 rz 180 deg; joints [-10.057, -79.362, 124.244, 165.892, 45.76, -133.526]
  MoveL 4619 to (-200, -41.2, 54.05) mm, rotated rx 128.92 ry 0 rz 180 deg; joints [-10.585, -78.775, 124.438, 165.357, 46.608, -130.908]
  MoveL 4620 to (0, -41.2, 54.05) mm, rotated rx 128.92 ry 0 rz 180 deg; joints [-9.07, -67.207, 108.731, 166.46, 42.326, -130.989]
  MoveL 4621 to (0, -40.82, 54.51) mm, rotated rx 131.3 ry 0 rz 180 deg; joints [-9.505, -66.699, 108.903, 166.005, 43.065, -128.377]
  MoveL 4622 to (-200, -40.82, 54.51) mm, rotated rx 131.3 ry 0 rz 180 deg; joints [-11.09, -78.16, 124.634, 164.873, 47.482, -128.343]
  MoveL 4623 to (-200, -40.41, 54.95) mm, rotated rx 133.69 ry 0 rz 180 deg; joints [-11.57, -77.515, 124.831, 164.438, 48.38, -125.83]
  MoveL 4624 to (0, -40.41, 54.95) mm, rotated rx 133.69 ry 0 rz 180 deg; joints [-9.919, -66.166, 109.076, 165.595, 43.823, -125.811]
  MoveL 4625 to (0, -39.99, 55.37) mm, rotated rx 136.08 ry 0 rz 180 deg; joints [-10.312, -65.612, 109.25, 165.229, 44.6, -123.29]
  MoveL 4626 to (-200, -39.99, 55.37) mm, rotated rx 136.08 ry 0 rz 180 deg; joints [-12.025, -76.843, 125.029, 164.05, 49.301, -123.366]
  MoveL 4627 to (-200, -39.55, 55.78) mm, rotated rx 138.47 ry 0 rz 180 deg; joints [-12.454, -76.144, 125.227, 163.708, 50.241, -120.947]
  MoveL 4628 to (0, -39.55, 55.78) mm, rotated rx 138.47 ry 0 rz 180 deg; joints [-10.684, -65.036, 109.424, 164.906, 45.394, -120.811]
  MoveL 4629 to (0, -39.09, 56.17) mm, rotated rx 140.85 ry 0 rz 180 deg; joints [-11.033, -64.438, 109.597, 164.625, 46.202, -118.373]
  MoveL 4630 to (-200, -39.09, 56.17) mm, rotated rx 140.85 ry 0 rz 180 deg; joints [-12.857, -75.419, 125.424, 163.409, 51.2, -118.573]
  MoveL 4631 to (-200, -38.62, 56.54) mm, rotated rx 143.24 ry 0 rz 180 deg; joints [-13.234, -74.669, 125.62, 163.153, 52.174, -116.241]
  MoveL 4632 to (0, -38.62, 56.54) mm, rotated rx 143.24 ry 0 rz 180 deg; joints [-11.359, -63.821, 109.769, 164.384, 47.024, -115.973]
  MoveL 4633 to (0, -38.13, 56.88) mm, rotated rx 145.63 ry 0 rz 180 deg; joints [-11.662, -63.185, 109.939, 164.18, 47.857, -113.608]
  MoveL 4634 to (-200, -38.13, 56.88) mm, rotated rx 145.63 ry 0 rz 180 deg; joints [-13.583, -73.895, 125.813, 162.936, 53.163, -113.945]
  MoveL 4635 to (-200, -37.63, 57.21) mm, rotated rx 148.01 ry 0 rz 180 deg; joints [-13.905, -73.099, 126.004, 162.757, 54.165, -111.687]
  MoveL 4636 to (0, -37.63, 57.21) mm, rotated rx 148.01 ry 0 rz 180 deg; joints [-11.941, -62.53, 110.107, 164.014, 48.7, -111.279]
  MoveL 4637 to (0, -37.11, 57.52) mm, rotated rx 150.4 ry 0 rz 180 deg; joints [-12.196, -61.858, 110.271, 163.882, 49.551, -108.981]
  MoveL 4638 to (-200, -37.11, 57.52) mm, rotated rx 150.4 ry 0 rz 180 deg; joints [-14.199, -72.28, 126.192, 162.615, 55.177, -109.462]
  MoveL 4639 to (-200, -36.59, 57.81) mm, rotated rx 152.79 ry 0 rz 180 deg; joints [-14.465, -71.441, 126.375, 162.507, 56.199, -107.266]
  MoveL 4640 to (0, -36.59, 57.81) mm, rotated rx 152.79 ry 0 rz 180 deg; joints [-12.427, -61.17, 110.433, 163.785, 50.409, -106.711]
  MoveL 4641 to (0, -36.05, 58.07) mm, rotated rx 155.18 ry 0 rz 180 deg; joints [-12.633, -60.466, 110.59, 163.719, 51.273, -104.47]
  MoveL 4642 to (-200, -36.05, 58.07) mm, rotated rx 155.18 ry 0 rz 180 deg; joints [-14.702, -70.583, 126.554, 162.432, 57.228, -105.1]
  MoveL 4643 to (-200, -35.5, 58.31) mm, rotated rx 157.56 ry 0 rz 180 deg; joints [-14.91, -69.707, 126.727, 162.389, 58.263, -102.958]
  MoveL 4644 to (0, -35.5, 58.31) mm, rotated rx 157.56 ry 0 rz 180 deg; joints [-12.814, -59.749, 110.743, 163.685, 52.141, -102.253]
  MoveL 4645 to (0, -34.94, 58.53) mm, rotated rx 159.95 ry 0 rz 180 deg; joints [-12.971, -59.018, 110.892, 163.68, 53.012, -100.058]
  MoveL 4646 to (-200, -34.94, 58.53) mm, rotated rx 159.95 ry 0 rz 180 deg; joints [-15.09, -68.814, 126.895, 162.377, 59.304, -100.838]
  MoveL 4647 to (-200, -34.37, 58.72) mm, rotated rx 162.34 ry 0 rz 180 deg; joints [-15.241, -67.906, 127.056, 162.393, 60.347, -98.739]
  MoveL 4648 to (0, -34.37, 58.72) mm, rotated rx 162.34 ry 0 rz 180 deg; joints [-13.102, -58.276, 111.035, 163.704, 53.885, -97.885]
  MoveL 4649 to (0, -33.79, 58.89) mm, rotated rx 164.72 ry 0 rz 180 deg; joints [-13.207, -57.523, 111.172, 163.755, 54.757, -95.73]
  MoveL 4650 to (-200, -33.79, 58.89) mm, rotated rx 164.72 ry 0 rz 180 deg; joints [-15.362, -66.984, 127.211, 162.437, 61.392, -96.657]
  MoveL 4651 to (-200, -33.21, 59.04) mm, rotated rx 167.11 ry 0 rz 180 deg; joints [-15.454, -66.049, 127.359, 162.507, 62.437, -94.59]
  MoveL 4652 to (0, -33.21, 59.04) mm, rotated rx 167.11 ry 0 rz 180 deg; joints [-13.288, -56.76, 111.304, 163.832, 55.629, -93.591]
  MoveL 4653 to (0, -32.62, 59.16) mm, rotated rx 169.5 ry 0 rz 180 deg; joints [-13.342, -55.99, 111.429, 163.934, 56.498, -91.468]
  MoveL 4654 to (-200, -32.62, 59.16) mm, rotated rx 169.5 ry 0 rz 180 deg; joints [-15.517, -65.104, 127.499, 162.604, 63.481, -92.537]
  MoveL 4655 to (-200, -32.03, 59.26) mm, rotated rx 171.89 ry 0 rz 180 deg; joints [-15.55, -64.15, 127.631, 162.725, 64.522, -90.494]
  MoveL 4656 to (0, -32.03, 59.26) mm, rotated rx 171.89 ry 0 rz 180 deg; joints [-13.371, -55.212, 111.548, 164.061, 57.364, -89.357]
  MoveL 4657 to (0, -31.44, 59.33) mm, rotated rx 174.28 ry 0 rz 180 deg; joints [-13.374, -54.429, 111.66, 164.212, 58.226, -87.257]
  MoveL 4658 to (-200, -31.44, 59.33) mm, rotated rx 174.28 ry 0 rz 180 deg; joints [-15.553, -63.188, 127.755, 162.871, 65.56, -88.458]
  MoveL 4659 to (-200, -30.84, 59.38) mm, rotated rx 176.66 ry 0 rz 180 deg; joints [-15.528, -62.221, 127.87, 163.04, 66.593, -86.43]
  MoveL 4660 to (0, -30.84, 59.38) mm, rotated rx 176.66 ry 0 rz 180 deg; joints [-13.352, -53.642, 111.765, 164.385, 59.082, -85.166]
  MoveL 4661 to (0, -30.24, 59.4) mm, rotated rx 179.05 ry 0 rz 180 deg; joints [-13.303, -52.852, 111.863, 164.58, 59.93, -83.083]
  MoveL 4662 to (-200, -30.24, 59.4) mm, rotated rx 179.05 ry 0 rz 180 deg; joints [-15.472, -61.249, 127.978, 163.232, 67.619, -84.406]
  MoveL 4663 to (-200, -29.64, 59.4) mm, rotated rx 180 ry 0 rz 180 deg; joints [-15.442, -60.838, 128.019, 163.317, 68.049, -83.608]
  MoveL 4664 to (0, -29.64, 59.4) mm, rotated rx 180 ry 0 rz 180 deg; joints [-13.277, -52.518, 111.902, 164.667, 60.286, -82.26]
  MoveL 4665 to (0, -29.04, 59.4) mm, rotated rx 180 ry 0 rz 180 deg; joints [-13.277, -52.486, 111.904, 164.672, 60.318, -82.271]
  MoveL 4666 to (-200, -29.04, 59.4) mm, rotated rx 180 ry 0 rz 180 deg; joints [-15.442, -60.799, 128.021, 163.322, 68.088, -83.62]
  MoveL 4667 to (-200, -28.44, 59.4) mm, rotated rx 180 ry 0 rz 180 deg; joints [-15.442, -60.761, 128.024, 163.326, 68.127, -83.633]
  MoveL 4668 to (0, -28.44, 59.4) mm, rotated rx 180 ry 0 rz 180 deg; joints [-13.277, -52.455, 111.906, 164.677, 60.35, -82.281]
  MoveL 4669 to (0, -27.84, 59.4) mm, rotated rx 180 ry 0 rz 180 deg; joints [-13.277, -52.424, 111.908, 164.682, 60.383, -82.291]
  MoveL 4670 to (-200, -27.84, 59.4) mm, rotated rx 180 ry 0 rz 180 deg; joints [-15.442, -60.722, 128.026, 163.331, 68.166, -83.646]
  MoveL 4671 to (-200, -27.24, 59.4) mm, rotated rx 180 ry 0 rz 180 deg; joints [-15.442, -60.684, 128.028, 163.336, 68.205, -83.658]
  MoveL 4672 to (0, -27.24, 59.4) mm, rotated rx 180 ry 0 rz 180 deg; joints [-13.277, -52.392, 111.91, 164.687, 60.415, -82.301]
  MoveL 4673 to (0, -26.64, 59.4) mm, rotated rx 180 ry 0 rz 180 deg; joints [-13.277, -52.361, 111.912, 164.692, 60.447, -82.311]
  MoveL 4674 to (-200, -26.64, 59.4) mm, rotated rx 180 ry 0 rz 180 deg; joints [-15.442, -60.645, 128.03, 163.34, 68.244, -83.671]
  MoveL 4675 to (-200, -26.04, 59.4) mm, rotated rx 180 ry 0 rz 180 deg; joints [-15.442, -60.607, 128.033, 163.345, 68.283, -83.683]
  MoveL 4676 to (0, -26.04, 59.4) mm, rotated rx 180 ry 0 rz 180 deg; joints [-13.277, -52.329, 111.914, 164.697, 60.479, -82.321]
  MoveL 4677 to (0, -25.44, 59.4) mm, rotated rx 180 ry 0 rz 180 deg; joints [-13.277, -52.298, 111.916, 164.702, 60.512, -82.332]
  MoveL 4678 to (-200, -25.44, 59.4) mm, rotated rx 180 ry 0 rz 180 deg; joints [-15.442, -60.568, 128.035, 163.35, 68.322, -83.696]
  MoveL 4679 to (-200, -24.84, 59.4) mm, rotated rx 180 ry 0 rz 180 deg; joints [-15.442, -60.529, 128.037, 163.354, 68.361, -83.709]
  MoveL 4680 to (0, -24.84, 59.4) mm, rotated rx 180 ry 0 rz 180 deg; joints [-13.277, -52.266, 111.918, 164.707, 60.544, -82.342]
  MoveL 4681 to (0, -24.24, 59.4) mm, rotated rx 180 ry 0 rz 180 deg; joints [-13.277, -52.235, 111.919, 164.712, 60.576, -82.352]
  MoveL 4682 to (-200, -24.24, 59.4) mm, rotated rx 180 ry 0 rz 180 deg; joints [-15.442, -60.491, 128.039, 163.359, 68.4, -83.721]
  MoveL 4683 to (-200, -23.64, 59.4) mm, rotated rx 180 ry 0 rz 180 deg; joints [-15.442, -60.452, 128.041, 163.364, 68.439, -83.734]
  MoveL 4684 to (0, -23.64, 59.4) mm, rotated rx 180 ry 0 rz 180 deg; joints [-13.277, -52.203, 111.921, 164.717, 60.608, -82.362]
  MoveL 4685 to (0, -23.04, 59.4) mm, rotated rx 180 ry 0 rz 180 deg; joints [-13.277, -52.172, 111.923, 164.722, 60.64, -82.372]
  MoveL 4686 to (-200, -23.04, 59.4) mm, rotated rx 180 ry 0 rz 180 deg; joints [-15.442, -60.414, 128.043, 163.368, 68.478, -83.746]
  MoveL 4687 to (-200, -22.44, 59.4) mm, rotated rx 180 ry 0 rz 180 deg; joints [-15.442, -60.375, 128.045, 163.373, 68.517, -83.759]
  MoveL 4688 to (0, -22.44, 59.4) mm, rotated rx 180 ry 0 rz 180 deg; joints [-13.277, -52.14, 111.925, 164.727, 60.672, -82.382]
  MoveL 4689 to (0, -21.84, 59.4) mm, rotated rx 180 ry 0 rz 180 deg; joints [-13.277, -52.109, 111.927, 164.732, 60.704, -82.392]
  MoveL 4690 to (-200, -21.84, 59.4) mm, rotated rx 180 ry 0 rz 180 deg; joints [-15.442, -60.336, 128.047, 163.377, 68.556, -83.771]
  MoveL 4691 to (-200, -21.24, 59.4) mm, rotated rx 180 ry 0 rz 180 deg; joints [-15.442, -60.297, 128.049, 163.382, 68.595, -83.784]
  MoveL 4692 to (0, -21.24, 59.4) mm, rotated rx 180 ry 0 rz 180 deg; joints [-13.277, -52.077, 111.928, 164.737, 60.737, -82.402]
  MoveL 4693 to (0, -20.64, 59.4) mm, rotated rx 180 ry 0 rz 180 deg; joints [-13.277, -52.046, 111.93, 164.742, 60.769, -82.412]
  MoveL 4694 to (-200, -20.64, 59.4) mm, rotated rx 180 ry 0 rz 180 deg; joints [-15.442, -60.259, 128.051, 163.387, 68.634, -83.796]
  MoveL 4695 to (-200, -20.04, 59.4) mm, rotated rx 180 ry 0 rz 180 deg; joints [-15.442, -60.22, 128.052, 163.391, 68.673, -83.809]
  MoveL 4696 to (0, -20.04, 59.4) mm, rotated rx 180 ry 0 rz 180 deg; joints [-13.277, -52.014, 111.932, 164.746, 60.801, -82.422]
  MoveL 4697 to (0, -19.44, 59.4) mm, rotated rx 180 ry 0 rz 180 deg; joints [-13.277, -51.982, 111.933, 164.751, 60.833, -82.432]
  MoveL 4698 to (-200, -19.44, 59.4) mm, rotated rx 180 ry 0 rz 180 deg; joints [-15.442, -60.181, 128.054, 163.396, 68.712, -83.821]
  MoveL 4699 to (-200, -18.84, 59.4) mm, rotated rx 180 ry 0 rz 180 deg; joints [-15.442, -60.142, 128.056, 163.4, 68.751, -83.833]
  MoveL 4700 to (0, -18.84, 59.4) mm, rotated rx 180 ry 0 rz 180 deg; joints [-13.277, -51.951, 111.935, 164.756, 60.865, -82.442]
  MoveL 4701 to (0, -18.24, 59.4) mm, rotated rx 180 ry 0 rz 180 deg; joints [-13.277, -51.919, 111.936, 164.761, 60.897, -82.452]
  MoveL 4702 to (-200, -18.24, 59.4) mm, rotated rx 180 ry 0 rz 180 deg; joints [-15.442, -60.104, 128.058, 163.405, 68.789, -83.846]
  MoveL 4703 to (-200, -17.64, 59.4) mm, rotated rx 180 ry 0 rz 180 deg; joints [-15.442, -60.065, 128.059, 163.409, 68.828, -83.858]
  MoveL 4704 to (0, -17.64, 59.4) mm, rotated rx 180 ry 0 rz 180 deg; joints [-13.277, -51.888, 111.938, 164.766, 60.929, -82.462]
  MoveL 4705 to (0, -17.04, 59.4) mm, rotated rx 180 ry 0 rz 180 deg; joints [-13.277, -51.856, 111.939, 164.771, 60.961, -82.472]
  MoveL 4706 to (-200, -17.04, 59.4) mm, rotated rx 180 ry 0 rz 180 deg; joints [-15.442, -60.026, 128.061, 163.414, 68.867, -83.871]
  MoveL 4707 to (-200, -16.44, 59.4) mm, rotated rx 180 ry 0 rz 180 deg; joints [-15.442, -59.987, 128.063, 163.418, 68.906, -83.883]
  MoveL 4708 to (0, -16.44, 59.4) mm, rotated rx 180 ry 0 rz 180 deg; joints [-13.277, -51.824, 111.941, 164.776, 60.993, -82.482]
  MoveL 4709 to (0, -15.84, 59.4) mm, rotated rx 180 ry 0 rz 180 deg; joints [-13.277, -51.792, 111.942, 164.78, 61.025, -82.492]
  MoveL 4710 to (-200, -15.84, 59.4) mm, rotated rx 180 ry 0 rz 180 deg; joints [-15.442, -59.948, 128.064, 163.422, 68.945, -83.895]
  MoveL 4711 to (-200, -15.24, 59.4) mm, rotated rx 180 ry 0 rz 180 deg; joints [-15.442, -59.909, 128.066, 163.427, 68.984, -83.908]
  MoveL 4712 to (0, -15.24, 59.4) mm, rotated rx 180 ry 0 rz 180 deg; joints [-13.277, -51.761, 111.944, 164.785, 61.057, -82.502]
  MoveL 4713 to (0, -14.64, 59.4) mm, rotated rx 180 ry 0 rz 180 deg; joints [-13.277, -51.729, 111.945, 164.79, 61.089, -82.512]
  MoveL 4714 to (-200, -14.64, 59.4) mm, rotated rx 180 ry 0 rz 180 deg; joints [-15.442, -59.87, 128.068, 163.431, 69.022, -83.92]
  MoveL 4715 to (-200, -14.04, 59.4) mm, rotated rx 180 ry 0 rz 180 deg; joints [-15.442, -59.831, 128.069, 163.436, 69.061, -83.933]
  MoveL 4716 to (0, -14.04, 59.4) mm, rotated rx 180 ry 0 rz 180 deg; joints [-13.277, -51.697, 111.947, 164.795, 61.121, -82.522]
  MoveL 4717 to (0, -13.44, 59.4) mm, rotated rx 180 ry 0 rz 180 deg; joints [-13.277, -51.665, 111.948, 164.8, 61.153, -82.532]
  MoveL 4718 to (-200, -13.44, 59.4) mm, rotated rx 180 ry 0 rz 180 deg; joints [-15.442, -59.792, 128.07, 163.44, 69.1, -83.945]
  MoveL 4719 to (-200, -12.84, 59.4) mm, rotated rx 180 ry 0 rz 180 deg; joints [-15.442, -59.753, 128.072, 163.445, 69.139, -83.957]
  MoveL 4720 to (0, -12.84, 59.4) mm, rotated rx 180 ry 0 rz 180 deg; joints [-13.277, -51.634, 111.949, 164.804, 61.185, -82.542]
  MoveL 4721 to (0, -12.24, 59.4) mm, rotated rx 180 ry 0 rz 180 deg; joints [-13.277, -51.602, 111.95, 164.809, 61.217, -82.552]
  MoveL 4722 to (-200, -12.24, 59.4) mm, rotated rx 180 ry 0 rz 180 deg; joints [-15.442, -59.714, 128.073, 163.449, 69.177, -83.97]
  MoveL 4723 to (-200, -11.64, 59.4) mm, rotated rx 180 ry 0 rz 180 deg; joints [-15.442, -59.675, 128.075, 163.453, 69.216, -83.982]
  MoveL 4724 to (0, -11.64, 59.4) mm, rotated rx 180 ry 0 rz 180 deg; joints [-13.277, -51.57, 111.952, 164.814, 61.249, -82.561]
  MoveL 4725 to (0, -11.04, 59.4) mm, rotated rx 180 ry 0 rz 180 deg; joints [-13.277, -51.538, 111.953, 164.819, 61.281, -82.571]
  MoveL 4726 to (-200, -11.04, 59.4) mm, rotated rx 180 ry 0 rz 180 deg; joints [-15.442, -59.636, 128.076, 163.458, 69.255, -83.994]
  MoveL 4727 to (-200, -10.44, 59.4) mm, rotated rx 180 ry 0 rz 180 deg; joints [-15.442, -59.597, 128.077, 163.462, 69.293, -84.006]
  MoveL 4728 to (0, -10.44, 59.4) mm, rotated rx 180 ry 0 rz 180 deg; joints [-13.277, -51.506, 111.954, 164.823, 61.312, -82.581]
  MoveL 4729 to (0, -9.84, 59.4) mm, rotated rx 180 ry 0 rz 180 deg; joints [-13.277, -51.474, 111.955, 164.828, 61.344, -82.591]
  MoveL 4730 to (-200, -9.84, 59.4) mm, rotated rx 180 ry 0 rz 180 deg; joints [-15.442, -59.558, 128.079, 163.466, 69.332, -84.019]
  MoveL 4731 to (-200, -9.24, 59.4) mm, rotated rx 180 ry 0 rz 180 deg; joints [-15.442, -59.519, 128.08, 163.471, 69.371, -84.031]
  MoveL 4732 to (0, -9.24, 59.4) mm, rotated rx 180 ry 0 rz 180 deg; joints [-13.277, -51.443, 111.956, 164.833, 61.376, -82.601]
  MoveL 4733 to (0, -8.64, 59.4) mm, rotated rx 180 ry 0 rz 180 deg; joints [-13.277, -51.411, 111.957, 164.838, 61.408, -82.611]
  MoveL 4734 to (-200, -8.64, 59.4) mm, rotated rx 180 ry 0 rz 180 deg; joints [-15.442, -59.48, 128.081, 163.475, 69.409, -84.043]
  MoveL 4735 to (-200, -8.04, 59.4) mm, rotated rx 180 ry 0 rz 180 deg; joints [-15.442, -59.441, 128.082, 163.479, 69.448, -84.055]
  MoveL 4736 to (0, -8.04, 59.4) mm, rotated rx 180 ry 0 rz 180 deg; joints [-13.277, -51.379, 111.959, 164.842, 61.44, -82.621]
  MoveL 4737 to (0, -7.44, 59.4) mm, rotated rx 180 ry 0 rz 180 deg; joints [-13.277, -51.347, 111.96, 164.847, 61.472, -82.63]
  MoveL 4738 to (-200, -7.44, 59.4) mm, rotated rx 180 ry 0 rz 180 deg; joints [-15.442, -59.402, 128.083, 163.484, 69.487, -84.068]
  MoveL 4739 to (-200, -6.84, 59.4) mm, rotated rx 180 ry 0 rz 180 deg; joints [-15.442, -59.363, 128.085, 163.488, 69.525, -84.08]
  MoveL 4740 to (0, -6.84, 59.4) mm, rotated rx 180 ry 0 rz 180 deg; joints [-13.277, -51.315, 111.961, 164.852, 61.503, -82.64]
  MoveL 4741 to (0, -6.24, 59.4) mm, rotated rx 180 ry 0 rz 180 deg; joints [-13.277, -51.283, 111.962, 164.856, 61.535, -82.65]
  MoveL 4742 to (-200, -6.24, 59.4) mm, rotated rx 180 ry 0 rz 180 deg; joints [-15.442, -59.323, 128.086, 163.492, 69.564, -84.092]
  MoveL 4743 to (-200, -5.64, 59.4) mm, rotated rx 180 ry 0 rz 180 deg; joints [-15.442, -59.284, 128.087, 163.496, 69.602, -84.104]
  MoveL 4744 to (0, -5.64, 59.4) mm, rotated rx 180 ry 0 rz 180 deg; joints [-13.277, -51.251, 111.962, 164.861, 61.567, -82.66]
  MoveL 4745 to (0, -5.04, 59.4) mm, rotated rx 180 ry 0 rz 180 deg; joints [-13.277, -51.219, 111.963, 164.866, 61.599, -82.669]
  MoveL 4746 to (-200, -5.04, 59.4) mm, rotated rx 180 ry 0 rz 180 deg; joints [-15.442, -59.245, 128.088, 163.501, 69.641, -84.116]
  MoveL 4747 to (-200, -4.44, 59.4) mm, rotated rx 180 ry 0 rz 180 deg; joints [-15.442, -59.206, 128.089, 163.505, 69.679, -84.129]
  MoveL 4748 to (0, -4.44, 59.4) mm, rotated rx 180 ry 0 rz 180 deg; joints [-13.277, -51.187, 111.964, 164.87, 61.63, -82.679]
  MoveL 4749 to (0, -3.84, 59.4) mm, rotated rx 180 ry 0 rz 180 deg; joints [-13.277, -51.155, 111.965, 164.875, 61.662, -82.689]
  MoveL 4750 to (-200, -3.84, 59.4) mm, rotated rx 180 ry 0 rz 180 deg; joints [-15.442, -59.167, 128.09, 163.509, 69.718, -84.141]
  MoveL 4751 to (-200, -3.24, 59.4) mm, rotated rx 180 ry 0 rz 180 deg; joints [-15.442, -59.127, 128.09, 163.513, 69.756, -84.153]
  MoveL 4752 to (0, -3.24, 59.4) mm, rotated rx 180 ry 0 rz 180 deg; joints [-13.277, -51.123, 111.966, 164.879, 61.694, -82.699]
  MoveL 4753 to (0, -2.64, 59.4) mm, rotated rx 180 ry 0 rz 180 deg; joints [-13.277, -51.091, 111.967, 164.884, 61.726, -82.708]
  MoveL 4754 to (-200, -2.64, 59.4) mm, rotated rx 180 ry 0 rz 180 deg; joints [-15.442, -59.088, 128.091, 163.517, 69.795, -84.165]
  MoveL 4755 to (-200, -2.04, 59.4) mm, rotated rx 180 ry 0 rz 180 deg; joints [-15.442, -59.049, 128.092, 163.522, 69.833, -84.177]
  MoveL 4756 to (0, -2.04, 59.4) mm, rotated rx 180 ry 0 rz 180 deg; joints [-13.277, -51.059, 111.967, 164.889, 61.757, -82.718]
  MoveL 4757 to (0, -1.44, 59.4) mm, rotated rx 180 ry 0 rz 180 deg; joints [-13.277, -51.027, 111.968, 164.893, 61.789, -82.728]
  MoveL 4758 to (-200, -1.44, 59.4) mm, rotated rx 180 ry 0 rz 180 deg; joints [-15.442, -59.01, 128.093, 163.526, 69.872, -84.189]
  MoveL 4759 to (-200, -0.84, 59.4) mm, rotated rx 180 ry 0 rz 180 deg; joints [-15.442, -58.97, 128.094, 163.53, 69.91, -84.201]
  MoveL 4760 to (0, -0.84, 59.4) mm, rotated rx 180 ry 0 rz 180 deg; joints [-13.277, -50.995, 111.969, 164.898, 61.821, -82.738]
  MoveL 4761 to (0, -0.24, 59.4) mm, rotated rx 180 ry 0 rz 180 deg; joints [-13.277, -50.962, 111.97, 164.902, 61.852, -82.747]
  MoveL 4762 to (-200, -0.24, 59.4) mm, rotated rx 180 ry 0 rz 180 deg; joints [-15.442, -58.931, 128.095, 163.534, 69.949, -84.214]
  MoveL 4763 to (-200, 0, 59.4) mm, rotated rx 180 ry 0 rz 180 deg; joints [-15.442, -58.915, 128.095, 163.536, 69.964, -84.218]
  MoveL 4764 to (0, 0, 59.4) mm, rotated rx 180 ry 0 rz 180 deg; joints [-13.277, -50.95, 111.97, 164.904, 61.865, -82.751]
  MoveL 4765 to (0, 0, 59.8) mm, rotated rx 180 ry 0 rz 180 deg; joints [-13.293, -50.946, 111.962, 164.886, 61.863, -82.741]
  MoveL 4766 to (-200, 0, 59.8) mm, rotated rx 180 ry 0 rz 180 deg; joints [-15.46, -58.911, 128.086, 163.516, 69.962, -84.21]
  MoveL 4767 to (-200, -0.6, 59.8) mm, rotated rx 180 ry 0 rz 180 deg; joints [-15.46, -58.95, 128.086, 163.512, 69.923, -84.198]
  MoveL 4768 to (0, -0.6, 59.8) mm, rotated rx 180 ry 0 rz 180 deg; joints [-13.293, -50.978, 111.961, 164.881, 61.831, -82.732]
  MoveL 4769 to (0, -1.2, 59.8) mm, rotated rx 180 ry 0 rz 180 deg; joints [-13.293, -51.01, 111.96, 164.877, 61.8, -82.722]
  MoveL 4770 to (-200, -1.2, 59.8) mm, rotated rx 180 ry 0 rz 180 deg; joints [-15.46, -58.99, 128.085, 163.508, 69.885, -84.186]
  MoveL 4771 to (-200, -1.8, 59.8) mm, rotated rx 180 ry 0 rz 180 deg; joints [-15.46, -59.029, 128.084, 163.504, 69.847, -84.174]
  MoveL 4772 to (0, -1.8, 59.8) mm, rotated rx 180 ry 0 rz 180 deg; joints [-13.293, -51.042, 111.96, 164.872, 61.768, -82.712]
  MoveL 4773 to (0, -2.4, 59.8) mm, rotated rx 180 ry 0 rz 180 deg; joints [-13.293, -51.074, 111.959, 164.868, 61.736, -82.703]
  MoveL 4774 to (-200, -2.4, 59.8) mm, rotated rx 180 ry 0 rz 180 deg; joints [-15.46, -59.068, 128.083, 163.499, 69.808, -84.162]
  MoveL 4775 to (-200, -3, 59.8) mm, rotated rx 180 ry 0 rz 180 deg; joints [-15.46, -59.108, 128.082, 163.495, 69.77, -84.15]
  MoveL 4776 to (0, -3, 59.8) mm, rotated rx 180 ry 0 rz 180 deg; joints [-13.293, -51.106, 111.958, 164.863, 61.705, -82.693]
  MoveL 4777 to (0, -3.6, 59.8) mm, rotated rx 180 ry 0 rz 180 deg; joints [-13.293, -51.138, 111.957, 164.858, 61.673, -82.683]
  MoveL 4778 to (-200, -3.6, 59.8) mm, rotated rx 180 ry 0 rz 180 deg; joints [-15.46, -59.147, 128.081, 163.491, 69.731, -84.138]
  MoveL 4779 to (-200, -4.2, 59.8) mm, rotated rx 180 ry 0 rz 180 deg; joints [-15.46, -59.186, 128.081, 163.487, 69.693, -84.126]
  MoveL 4780 to (0, -4.2, 59.8) mm, rotated rx 180 ry 0 rz 180 deg; joints [-13.293, -51.17, 111.957, 164.854, 61.641, -82.673]
  MoveL 4781 to (0, -4.8, 59.8) mm, rotated rx 180 ry 0 rz 180 deg; joints [-13.293, -51.202, 111.956, 164.849, 61.61, -82.664]
  MoveL 4782 to (-200, -4.8, 59.8) mm, rotated rx 180 ry 0 rz 180 deg; joints [-15.46, -59.225, 128.08, 163.483, 69.654, -84.113]
  MoveL 4783 to (-200, -5.4, 59.8) mm, rotated rx 180 ry 0 rz 180 deg; joints [-15.46, -59.264, 128.079, 163.478, 69.616, -84.101]
  MoveL 4784 to (0, -5.4, 59.8) mm, rotated rx 180 ry 0 rz 180 deg; joints [-13.293, -51.234, 111.955, 164.844, 61.578, -82.654]
  MoveL 4785 to (0, -6, 59.8) mm, rotated rx 180 ry 0 rz 180 deg; joints [-13.293, -51.266, 111.954, 164.84, 61.546, -82.644]
  MoveL 4786 to (-200, -6, 59.8) mm, rotated rx 180 ry 0 rz 180 deg; joints [-15.46, -59.304, 128.078, 163.474, 69.577, -84.089]
  MoveL 4787 to (-200, -6.6, 59.8) mm, rotated rx 180 ry 0 rz 180 deg; joints [-15.46, -59.343, 128.076, 163.47, 69.538, -84.077]
  MoveL 4788 to (0, -6.6, 59.8) mm, rotated rx 180 ry 0 rz 180 deg; joints [-13.293, -51.298, 111.953, 164.835, 61.514, -82.634]
  MoveL 4789 to (0, -7.2, 59.8) mm, rotated rx 180 ry 0 rz 180 deg; joints [-13.293, -51.33, 111.952, 164.83, 61.482, -82.624]
  MoveL 4790 to (-200, -7.2, 59.8) mm, rotated rx 180 ry 0 rz 180 deg; joints [-15.46, -59.382, 128.075, 163.466, 69.5, -84.064]
  MoveL 4791 to (-200, -7.8, 59.8) mm, rotated rx 180 ry 0 rz 180 deg; joints [-15.46, -59.421, 128.074, 163.461, 69.461, -84.052]
  MoveL 4792 to (0, -7.8, 59.8) mm, rotated rx 180 ry 0 rz 180 deg; joints [-13.293, -51.362, 111.951, 164.826, 61.451, -82.615]
  MoveL 4793 to (0, -8.4, 59.8) mm, rotated rx 180 ry 0 rz 180 deg; joints [-13.293, -51.394, 111.95, 164.821, 61.419, -82.605]
  MoveL 4794 to (-200, -8.4, 59.8) mm, rotated rx 180 ry 0 rz 180 deg; joints [-15.46, -59.46, 128.073, 163.457, 69.423, -84.04]
  MoveL 4795 to (-200, -9, 59.8) mm, rotated rx 180 ry 0 rz 180 deg; joints [-15.46, -59.499, 128.072, 163.453, 69.384, -84.028]
  MoveL 4796 to (0, -9, 59.8) mm, rotated rx 180 ry 0 rz 180 deg; joints [-13.293, -51.426, 111.949, 164.816, 61.387, -82.595]
  MoveL 4797 to (0, -9.6, 59.8) mm, rotated rx 180 ry 0 rz 180 deg; joints [-13.293, -51.458, 111.948, 164.812, 61.355, -82.585]
  MoveL 4798 to (-200, -9.6, 59.8) mm, rotated rx 180 ry 0 rz 180 deg; joints [-15.46, -59.538, 128.071, 163.448, 69.345, -84.015]
  MoveL 4799 to (-200, -10.2, 59.8) mm, rotated rx 180 ry 0 rz 180 deg; joints [-15.46, -59.577, 128.069, 163.444, 69.307, -84.003]
  MoveL 4800 to (0, -10.2, 59.8) mm, rotated rx 180 ry 0 rz 180 deg; joints [-13.293, -51.49, 111.946, 164.807, 61.323, -82.575]
  MoveL 4801 to (0, -10.8, 59.8) mm, rotated rx 180 ry 0 rz 180 deg; joints [-13.293, -51.521, 111.945, 164.802, 61.291, -82.565]
  MoveL 4802 to (-200, -10.8, 59.8) mm, rotated rx 180 ry 0 rz 180 deg; joints [-15.46, -59.617, 128.068, 163.44, 69.268, -83.991]
  MoveL 4803 to (-200, -11.4, 59.8) mm, rotated rx 180 ry 0 rz 180 deg; joints [-15.46, -59.656, 128.067, 163.435, 69.229, -83.979]
  MoveL 4804 to (0, -11.4, 59.8) mm, rotated rx 180 ry 0 rz 180 deg; joints [-13.293, -51.553, 111.944, 164.797, 61.26, -82.556]
  MoveL 4805 to (0, -12, 59.8) mm, rotated rx 180 ry 0 rz 180 deg; joints [-13.293, -51.585, 111.943, 164.793, 61.228, -82.546]
  MoveL 4806 to (-200, -12, 59.8) mm, rotated rx 180 ry 0 rz 180 deg; joints [-15.46, -59.695, 128.065, 163.431, 69.191, -83.966]
  MoveL 4807 to (-200, -12.6, 59.8) mm, rotated rx 180 ry 0 rz 180 deg; joints [-15.46, -59.734, 128.064, 163.427, 69.152, -83.954]
  MoveL 4808 to (0, -12.6, 59.8) mm, rotated rx 180 ry 0 rz 180 deg; joints [-13.293, -51.617, 111.942, 164.788, 61.196, -82.536]
  MoveL 4809 to (0, -13.2, 59.8) mm, rotated rx 180 ry 0 rz 180 deg; joints [-13.293, -51.649, 111.94, 164.783, 61.164, -82.526]
  MoveL 4810 to (-200, -13.2, 59.8) mm, rotated rx 180 ry 0 rz 180 deg; joints [-15.46, -59.773, 128.063, 163.422, 69.113, -83.942]
  MoveL 4811 to (-200, -13.8, 59.8) mm, rotated rx 180 ry 0 rz 180 deg; joints [-15.46, -59.811, 128.061, 163.418, 69.074, -83.929]
  MoveL 4812 to (0, -13.8, 59.8) mm, rotated rx 180 ry 0 rz 180 deg; joints [-13.293, -51.68, 111.939, 164.778, 61.132, -82.516]
  MoveL 4813 to (0, -14.4, 59.8) mm, rotated rx 180 ry 0 rz 180 deg; joints [-13.293, -51.712, 111.938, 164.773, 61.1, -82.506]
  MoveL 4814 to (-200, -14.4, 59.8) mm, rotated rx 180 ry 0 rz 180 deg; joints [-15.46, -59.85, 128.06, 163.413, 69.036, -83.917]
  MoveL 4815 to (-200, -15, 59.8) mm, rotated rx 180 ry 0 rz 180 deg; joints [-15.46, -59.889, 128.058, 163.409, 68.997, -83.905]
  MoveL 4816 to (0, -15, 59.8) mm, rotated rx 180 ry 0 rz 180 deg; joints [-13.293, -51.744, 111.936, 164.769, 61.068, -82.496]
  MoveL 4817 to (0, -15.6, 59.8) mm, rotated rx 180 ry 0 rz 180 deg; joints [-13.293, -51.776, 111.935, 164.764, 61.036, -82.486]
  MoveL 4818 to (-200, -15.6, 59.8) mm, rotated rx 180 ry 0 rz 180 deg; joints [-15.46, -59.928, 128.057, 163.404, 68.958, -83.892]
  MoveL 4819 to (-200, -16.2, 59.8) mm, rotated rx 180 ry 0 rz 180 deg; joints [-15.46, -59.967, 128.055, 163.4, 68.919, -83.88]
  MoveL 4820 to (0, -16.2, 59.8) mm, rotated rx 180 ry 0 rz 180 deg; joints [-13.293, -51.807, 111.933, 164.759, 61.004, -82.476]
  MoveL 4821 to (0, -16.8, 59.8) mm, rotated rx 180 ry 0 rz 180 deg; joints [-13.293, -51.839, 111.932, 164.754, 60.972, -82.466]
  MoveL 4822 to (-200, -16.8, 59.8) mm, rotated rx 180 ry 0 rz 180 deg; joints [-15.46, -60.006, 128.053, 163.396, 68.881, -83.867]
  MoveL 4823 to (-200, -17.4, 59.8) mm, rotated rx 180 ry 0 rz 180 deg; joints [-15.46, -60.045, 128.052, 163.391, 68.842, -83.855]
  MoveL 4824 to (0, -17.4, 59.8) mm, rotated rx 180 ry 0 rz 180 deg; joints [-13.293, -51.871, 111.931, 164.749, 60.94, -82.456]
  MoveL 4825 to (0, -18, 59.8) mm, rotated rx 180 ry 0 rz 180 deg; joints [-13.293, -51.902, 111.929, 164.744, 60.908, -82.446]
  MoveL 4826 to (-200, -18, 59.8) mm, rotated rx 180 ry 0 rz 180 deg; joints [-15.46, -60.084, 128.05, 163.387, 68.803, -83.843]
  MoveL 4827 to (-200, -18.6, 59.8) mm, rotated rx 180 ry 0 rz 180 deg; joints [-15.46, -60.123, 128.048, 163.382, 68.764, -83.83]
  MoveL 4828 to (0, -18.6, 59.8) mm, rotated rx 180 ry 0 rz 180 deg; joints [-13.293, -51.934, 111.927, 164.74, 60.876, -82.436]
  MoveL 4829 to (0, -19.2, 59.8) mm, rotated rx 180 ry 0 rz 180 deg; joints [-13.293, -51.966, 111.926, 164.735, 60.844, -82.426]
  MoveL 4830 to (-200, -19.2, 59.8) mm, rotated rx 180 ry 0 rz 180 deg; joints [-15.46, -60.161, 128.047, 163.378, 68.725, -83.818]
  MoveL 4831 to (-200, -19.8, 59.8) mm, rotated rx 180 ry 0 rz 180 deg; joints [-15.46, -60.2, 128.045, 163.373, 68.686, -83.805]
  MoveL 4832 to (0, -19.8, 59.8) mm, rotated rx 180 ry 0 rz 180 deg; joints [-13.293, -51.997, 111.924, 164.73, 60.812, -82.416]
  MoveL 4833 to (0, -20.4, 59.8) mm, rotated rx 180 ry 0 rz 180 deg; joints [-13.293, -52.029, 111.923, 164.725, 60.78, -82.406]
  MoveL 4834 to (-200, -20.4, 59.8) mm, rotated rx 180 ry 0 rz 180 deg; joints [-15.46, -60.239, 128.043, 163.368, 68.647, -83.793]
  MoveL 4835 to (-200, -21, 59.8) mm, rotated rx 180 ry 0 rz 180 deg; joints [-15.46, -60.278, 128.041, 163.364, 68.609, -83.78]
  MoveL 4836 to (0, -21, 59.8) mm, rotated rx 180 ry 0 rz 180 deg; joints [-13.293, -52.061, 111.921, 164.72, 60.748, -82.396]
  MoveL 4837 to (0, -21.6, 59.8) mm, rotated rx 180 ry 0 rz 180 deg; joints [-13.293, -52.092, 111.919, 164.715, 60.716, -82.386]
  MoveL 4838 to (-200, -21.6, 59.8) mm, rotated rx 180 ry 0 rz 180 deg; joints [-15.46, -60.316, 128.039, 163.359, 68.57, -83.768]
  MoveL 4839 to (-200, -22.2, 59.8) mm, rotated rx 180 ry 0 rz 180 deg; joints [-15.46, -60.355, 128.037, 163.355, 68.531, -83.755]
  MoveL 4840 to (0, -22.2, 59.8) mm, rotated rx 180 ry 0 rz 180 deg; joints [-13.293, -52.124, 111.917, 164.71, 60.683, -82.376]
  MoveL 4841 to (0, -22.8, 59.8) mm, rotated rx 180 ry 0 rz 180 deg; joints [-13.293, -52.155, 111.916, 164.705, 60.651, -82.366]
  MoveL 4842 to (-200, -22.8, 59.8) mm, rotated rx 180 ry 0 rz 180 deg; joints [-15.46, -60.394, 128.035, 163.35, 68.492, -83.743]
  MoveL 4843 to (-200, -23.4, 59.8) mm, rotated rx 180 ry 0 rz 180 deg; joints [-15.46, -60.432, 128.033, 163.346, 68.453, -83.73]
  MoveL 4844 to (0, -23.4, 59.8) mm, rotated rx 180 ry 0 rz 180 deg; joints [-13.293, -52.187, 111.914, 164.7, 60.619, -82.356]
  MoveL 4845 to (0, -24, 59.8) mm, rotated rx 180 ry 0 rz 180 deg; joints [-13.293, -52.218, 111.912, 164.695, 60.587, -82.346]
  MoveL 4846 to (-200, -24, 59.8) mm, rotated rx 180 ry 0 rz 180 deg; joints [-15.46, -60.471, 128.031, 163.341, 68.414, -83.718]
  MoveL 4847 to (-200, -24.6, 59.8) mm, rotated rx 180 ry 0 rz 180 deg; joints [-15.46, -60.51, 128.029, 163.336, 68.375, -83.705]
  MoveL 4848 to (0, -24.6, 59.8) mm, rotated rx 180 ry 0 rz 180 deg; joints [-13.293, -52.25, 111.91, 164.69, 60.555, -82.336]
  MoveL 4849 to (0, -25.2, 59.8) mm, rotated rx 180 ry 0 rz 180 deg; joints [-13.293, -52.281, 111.908, 164.685, 60.523, -82.325]
  MoveL 4850 to (-200, -25.2, 59.8) mm, rotated rx 180 ry 0 rz 180 deg; joints [-15.46, -60.548, 128.027, 163.332, 68.336, -83.693]
  MoveL 4851 to (-200, -25.8, 59.8) mm, rotated rx 180 ry 0 rz 180 deg; joints [-15.46, -60.587, 128.025, 163.327, 68.297, -83.68]
  MoveL 4852 to (0, -25.8, 59.8) mm, rotated rx 180 ry 0 rz 180 deg; joints [-13.293, -52.313, 111.906, 164.68, 60.49, -82.315]
  MoveL 4853 to (0, -26.4, 59.8) mm, rotated rx 180 ry 0 rz 180 deg; joints [-13.293, -52.344, 111.905, 164.675, 60.458, -82.305]
  MoveL 4854 to (-200, -26.4, 59.8) mm, rotated rx 180 ry 0 rz 180 deg; joints [-15.46, -60.626, 128.023, 163.322, 68.258, -83.667]
  MoveL 4855 to (-200, -27, 59.8) mm, rotated rx 180 ry 0 rz 180 deg; joints [-15.46, -60.664, 128.021, 163.318, 68.219, -83.655]
  MoveL 4856 to (0, -27, 59.8) mm, rotated rx 180 ry 0 rz 180 deg; joints [-13.293, -52.376, 111.903, 164.67, 60.426, -82.295]
  MoveL 4857 to (0, -27.6, 59.8) mm, rotated rx 180 ry 0 rz 180 deg; joints [-13.293, -52.407, 111.901, 164.665, 60.394, -82.285]
  MoveL 4858 to (-200, -27.6, 59.8) mm, rotated rx 180 ry 0 rz 180 deg; joints [-15.46, -60.703, 128.018, 163.313, 68.18, -83.642]
  MoveL 4859 to (-200, -28.2, 59.8) mm, rotated rx 180 ry 0 rz 180 deg; joints [-15.46, -60.741, 128.016, 163.308, 68.141, -83.63]
  MoveL 4860 to (0, -28.2, 59.8) mm, rotated rx 180 ry 0 rz 180 deg; joints [-13.293, -52.438, 111.899, 164.66, 60.362, -82.275]
  MoveL 4861 to (0, -28.8, 59.8) mm, rotated rx 180 ry 0 rz 180 deg; joints [-13.293, -52.47, 111.896, 164.655, 60.329, -82.265]
  MoveL 4862 to (-200, -28.8, 59.8) mm, rotated rx 180 ry 0 rz 180 deg; joints [-15.46, -60.78, 128.014, 163.304, 68.102, -83.617]
  MoveL 4863 to (-200, -29.4, 59.8) mm, rotated rx 180 ry 0 rz 180 deg; joints [-15.46, -60.818, 128.012, 163.299, 68.062, -83.604]
  MoveL 4864 to (0, -29.4, 59.8) mm, rotated rx 180 ry 0 rz 180 deg; joints [-13.293, -52.501, 111.894, 164.65, 60.297, -82.254]
  MoveL 4865 to (0, -30, 59.8) mm, rotated rx 180 ry 0 rz 180 deg; joints [-13.293, -52.533, 111.892, 164.645, 60.265, -82.244]
  MoveL 4866 to (-200, -30, 59.8) mm, rotated rx 180 ry 0 rz 180 deg; joints [-15.46, -60.857, 128.009, 163.294, 68.023, -83.592]
  MoveL 4867 to (-200, -30.6, 59.79) mm, rotated rx 177.68 ry 0 rz 180 deg; joints [-15.526, -61.804, 127.908, 163.098, 67.027, -85.56]
  MoveL 4868 to (0, -30.6, 59.79) mm, rotated rx 177.68 ry 0 rz 180 deg; joints [-13.35, -53.303, 111.8, 164.446, 59.441, -84.268]
  MoveL 4869 to (0, -31.2, 59.75) mm, rotated rx 175.35 ry 0 rz 180 deg; joints [-13.383, -54.071, 111.7, 164.268, 58.61, -86.299]
  MoveL 4870 to (-200, -31.2, 59.75) mm, rotated rx 175.35 ry 0 rz 180 deg; joints [-15.564, -62.749, 127.799, 162.924, 66.024, -87.531]
  MoveL 4871 to (-200, -31.8, 59.69) mm, rotated rx 173.03 ry 0 rz 180 deg; joints [-15.573, -63.688, 127.682, 162.771, 65.016, -89.506]
  MoveL 4872 to (0, -31.8, 59.69) mm, rotated rx 173.03 ry 0 rz 180 deg; joints [-13.391, -54.835, 111.594, 164.111, 57.774, -88.337]
  MoveL 4873 to (0, -32.39, 59.61) mm, rotated rx 170.71 ry 0 rz 180 deg; joints [-13.376, -55.595, 111.482, 163.976, 56.933, -90.385]
  MoveL 4874 to (-200, -32.39, 59.61) mm, rotated rx 170.71 ry 0 rz 180 deg; joints [-15.555, -64.621, 127.558, 162.641, 64.004, -91.489]
  MoveL 4875 to (-200, -32.98, 59.5) mm, rotated rx 168.39 ry 0 rz 180 deg; joints [-15.509, -65.546, 127.425, 162.535, 62.988, -93.481]
  MoveL 4876 to (0, -32.98, 59.5) mm, rotated rx 168.39 ry 0 rz 180 deg; joints [-13.335, -56.35, 111.363, 163.863, 56.088, -92.444]
  MoveL 4877 to (0, -33.56, 59.36) mm, rotated rx 166.06 ry 0 rz 180 deg; joints [-13.271, -57.097, 111.238, 163.775, 55.24, -94.516]
  MoveL 4878 to (-200, -33.56, 59.36) mm, rotated rx 166.06 ry 0 rz 180 deg; joints [-15.435, -66.462, 127.285, 162.452, 61.97, -95.485]
  MoveL 4879 to (-200, -34.14, 59.21) mm, rotated rx 163.74 ry 0 rz 180 deg; joints [-15.333, -67.367, 127.138, 162.394, 60.953, -97.501]
  MoveL 4880 to (0, -34.14, 59.21) mm, rotated rx 163.74 ry 0 rz 180 deg; joints [-13.182, -57.836, 111.107, 163.71, 54.39, -96.603]
  MoveL 4881 to (0, -34.72, 59.03) mm, rotated rx 161.42 ry 0 rz 180 deg; joints [-13.069, -58.565, 110.971, 163.671, 53.541, -98.706]
  MoveL 4882 to (-200, -34.72, 59.03) mm, rotated rx 161.42 ry 0 rz 180 deg; joints [-15.203, -68.26, 126.985, 162.361, 59.936, -99.531]
  MoveL 4883 to (-200, -35.28, 58.83) mm, rotated rx 159.09 ry 0 rz 180 deg; joints [-15.046, -69.139, 126.825, 162.356, 58.921, -101.581]
  MoveL 4884 to (0, -35.28, 58.83) mm, rotated rx 159.09 ry 0 rz 180 deg; joints [-12.932, -59.284, 110.83, 163.658, 52.691, -100.827]
  MoveL 4885 to (0, -35.84, 58.6) mm, rotated rx 156.77 ry 0 rz 180 deg; joints [-12.772, -59.991, 110.684, 163.672, 51.844, -102.969]
  MoveL 4886 to (-200, -35.84, 58.6) mm, rotated rx 156.77 ry 0 rz 180 deg; joints [-14.861, -70.003, 126.66, 162.378, 57.909, -103.65]
  MoveL 4887 to (-200, -36.38, 58.35) mm, rotated rx 154.45 ry 0 rz 180 deg; joints [-14.649, -70.851, 126.489, 162.429, 56.903, -105.741]
  MoveL 4888 to (0, -36.38, 58.35) mm, rotated rx 154.45 ry 0 rz 180 deg; joints [-12.587, -60.685, 110.533, 163.715, 51, -105.133]
  MoveL 4889 to (0, -36.92, 58.08) mm, rotated rx 152.13 ry 0 rz 180 deg; joints [-12.379, -61.366, 110.378, 163.787, 50.16, -107.322]
  MoveL 4890 to (-200, -36.92, 58.08) mm, rotated rx 152.13 ry 0 rz 180 deg; joints [-14.41, -71.681, 126.314, 162.511, 55.902, -107.857]
  MoveL 4891 to (-200, -37.44, 57.79) mm, rotated rx 149.8 ry 0 rz 180 deg; joints [-14.144, -72.493, 126.134, 162.624, 54.91, -109.998]
  MoveL 4892 to (0, -37.44, 57.79) mm, rotated rx 149.8 ry 0 rz 180 deg; joints [-12.148, -62.032, 110.22, 163.891, 49.326, -109.536]
  MoveL 4893 to (0, -37.96, 57.48) mm, rotated rx 147.48 ry 0 rz 180 deg; joints [-11.894, -62.683, 110.059, 164.026, 48.498, -111.779]
  MoveL 4894 to (-200, -37.96, 57.48) mm, rotated rx 147.48 ry 0 rz 180 deg; joints [-13.851, -73.285, 125.951, 162.771, 53.926, -112.171]
  MoveL 4895 to (-200, -38.45, 57.15) mm, rotated rx 145.16 ry 0 rz 180 deg; joints [-13.532, -74.056, 125.764, 162.953, 52.953, -114.375]
  MoveL 4896 to (0, -38.45, 57.15) mm, rotated rx 145.16 ry 0 rz 180 deg; joints [-11.617, -63.317, 109.895, 164.196, 47.679, -114.052]
  MoveL 4897 to (0, -38.94, 56.79) mm, rotated rx 142.84 ry 0 rz 180 deg; joints [-11.318, -63.933, 109.729, 164.4, 46.87, -116.358]
  MoveL 4898 to (-200, -38.94, 56.79) mm, rotated rx 142.84 ry 0 rz 180 deg; joints [-13.187, -74.806, 125.575, 163.171, 51.992, -116.614]
  MoveL 4899 to (-200, -39.41, 56.42) mm, rotated rx 140.51 ry 0 rz 180 deg; joints [-12.816, -75.532, 125.384, 163.427, 51.046, -118.89]
  MoveL 4900 to (0, -39.41, 56.42) mm, rotated rx 140.51 ry 0 rz 180 deg; joints [-10.997, -64.531, 109.561, 164.641, 46.071, -118.699]
  MoveL 4901 to (0, -39.87, 56.03) mm, rotated rx 138.19 ry 0 rz 180 deg; joints [-10.654, -65.11, 109.393, 164.92, 45.286, -121.076]
  MoveL 4902 to (-200, -39.87, 56.03) mm, rotated rx 138.19 ry 0 rz 180 deg; joints [-12.42, -76.235, 125.192, 163.722, 50.114, -121.204]
  MoveL 4903 to (-200, -40.31, 55.62) mm, rotated rx 135.87 ry 0 rz 180 deg; joints [-11.999, -76.913, 124.999, 164.06, 49.2, -123.562]
  MoveL 4904 to (0, -40.31, 55.62) mm, rotated rx 135.87 ry 0 rz 180 deg; joints [-10.29, -65.669, 109.223, 165.238, 44.515, -123.492]
  MoveL 4905 to (0, -40.73, 55.2) mm, rotated rx 133.54 ry 0 rz 180 deg; joints [-9.906, -66.208, 109.054, 165.598, 43.759, -125.948]
  MoveL 4906 to (-200, -40.73, 55.2) mm, rotated rx 133.54 ry 0 rz 180 deg; joints [-11.554, -77.565, 124.806, 164.441, 48.305, -125.963]
  MoveL 4907 to (-200, -41.13, 54.75) mm, rotated rx 131.22 ry 0 rz 180 deg; joints [-11.085, -78.191, 124.614, 164.866, 47.432, -128.411]
  MoveL 4908 to (0, -41.13, 54.75) mm, rotated rx 131.22 ry 0 rz 180 deg; joints [-9.501, -66.725, 108.885, 165.999, 43.021, -128.448]
  MoveL 4909 to (0, -41.52, 54.29) mm, rotated rx 128.9 ry 0 rz 180 deg; joints [-9.077, -67.22, 108.717, 166.444, 42.302, -130.991]
  MoveL 4910 to (-200, -41.52, 54.29) mm, rotated rx 128.9 ry 0 rz 180 deg; joints [-10.593, -78.791, 124.424, 165.339, 46.581, -130.908]
  MoveL 4911 to (-200, -41.88, 53.82) mm, rotated rx 126.58 ry 0 rz 180 deg; joints [-10.079, -79.361, 124.235, 165.859, 45.755, -133.454]
  MoveL 4912 to (0, -41.88, 53.82) mm, rotated rx 126.58 ry 0 rz 180 deg; joints [-8.634, -67.692, 108.552, 166.933, 41.605, -133.578]
  MoveL 4913 to (0, -42.23, 53.33) mm, rotated rx 124.25 ry 0 rz 180 deg; joints [-8.173, -68.141, 108.388, 167.468, 40.929, -136.214]
  MoveL 4914 to (-200, -42.23, 53.33) mm, rotated rx 124.25 ry 0 rz 180 deg; joints [-9.543, -79.904, 124.049, 166.429, 44.956, -136.053]
  MoveL 4915 to (-200, -42.56, 52.83) mm, rotated rx 121.93 ry 0 rz 180 deg; joints [-8.986, -80.418, 123.866, 167.05, 44.186, -138.706]
  MoveL 4916 to (0, -42.56, 52.83) mm, rotated rx 121.93 ry 0 rz 180 deg; joints [-7.693, -68.567, 108.227, 168.049, 40.278, -138.897]
  MoveL 4917 to (0, -42.87, 52.31) mm, rotated rx 119.61 ry 0 rz 180 deg; joints [-7.198, -68.967, 108.069, 168.677, 39.654, -141.629]
  MoveL 4918 to (-200, -42.87, 52.31) mm, rotated rx 119.61 ry 0 rz 180 deg; joints [-8.409, -80.901, 123.688, 167.722, 43.448, -141.414]
  MoveL 4919 to (-200, -43.15, 51.78) mm, rotated rx 117.28 ry 0 rz 180 deg; joints [-7.813, -81.355, 123.514, 168.446, 42.743, -144.177]
  MoveL 4920 to (0, -43.15, 51.78) mm, rotated rx 117.28 ry 0 rz 180 deg; joints [-6.685, -69.344, 107.916, 169.353, 39.058, -144.411]
  MoveL 4921 to (0, -43.42, 51.25) mm, rotated rx 114.96 ry 0 rz 180 deg; joints [-6.158, -69.694, 107.766, 170.075, 38.492, -147.24]
  MoveL 4922 to (-200, -43.42, 51.25) mm, rotated rx 114.96 ry 0 rz 180 deg; joints [-7.199, -81.778, 123.345, 169.221, 42.075, -146.995]
  MoveL 4923 to (-200, -43.66, 50.7) mm, rotated rx 112.64 ry 0 rz 180 deg; joints [-6.567, -82.169, 123.183, 170.049, 41.444, -149.869]
  MoveL 4924 to (0, -43.66, 50.7) mm, rotated rx 112.64 ry 0 rz 180 deg; joints [-5.617, -70.019, 107.622, 170.844, 37.958, -150.119]
  MoveL 4925 to (0, -43.88, 50.14) mm, rotated rx 110.32 ry 0 rz 180 deg; joints [-5.062, -70.318, 107.483, 171.659, 37.458, -153.046]
  MoveL 4926 to (-200, -43.88, 50.14) mm, rotated rx 110.32 ry 0 rz 180 deg; joints [-5.92, -82.529, 123.026, 170.929, 40.854, -152.798]
  MoveL 4927 to (-200, -44.08, 49.57) mm, rotated rx 107.99 ry 0 rz 180 deg; joints [-5.257, -82.857, 122.877, 171.858, 40.307, -155.78]
  MoveL 4928 to (0, -44.08, 49.57) mm, rotated rx 107.99 ry 0 rz 180 deg; joints [-4.494, -70.591, 107.35, 172.518, 36.994, -156.019]
  MoveL 4929 to (0, -44.25, 49) mm, rotated rx 105.67 ry 0 rz 180 deg; joints [-3.915, -70.837, 107.223, 173.42, 36.567, -159.037]
  MoveL 4930 to (-200, -44.25, 49) mm, rotated rx 105.67 ry 0 rz 180 deg; joints [-4.58, -83.152, 122.735, 172.835, 39.804, -158.813]
  MoveL 4931 to (-200, -44.4, 48.42) mm, rotated rx 103.35 ry 0 rz 180 deg; joints [-3.891, -83.415, 122.602, 173.856, 39.349, -161.894]
  MoveL 4932 to (0, -44.4, 48.42) mm, rotated rx 103.35 ry 0 rz 180 deg; joints [-3.325, -71.056, 107.103, 174.362, 36.18, -162.096]
  MoveL 4933 to (0, -44.53, 47.83) mm, rotated rx 101.03 ry 0 rz 180 deg; joints [-2.726, -71.247, 106.99, 175.341, 35.833, -165.195]
  MoveL 4934 to (-200, -44.53, 47.83) mm, rotated rx 101.03 ry 0 rz 180 deg; joints [-3.19, -83.645, 122.477, 174.921, 38.942, -165.02]
  MoveL 4935 to (-200, -44.63, 47.24) mm, rotated rx 98.7 ry 0 rz 180 deg; joints [-2.479, -83.842, 122.36, 176.023, 38.586, -168.187]
  MoveL 4936 to (0, -44.63, 47.24) mm, rotated rx 98.7 ry 0 rz 180 deg; joints [-2.118, -71.411, 106.885, 176.353, 35.528, -168.329]
  MoveL 4937 to (0, -44.71, 46.64) mm, rotated rx 96.38 ry 0 rz 180 deg; joints [-1.503, -71.548, 106.787, 177.396, 35.267, -171.495]
  MoveL 4938 to (-200, -44.71, 46.64) mm, rotated rx 96.38 ry 0 rz 180 deg; joints [-1.76, -84.005, 122.253, 177.159, 38.282, -171.39]
  MoveL 4939 to (-200, -44.76, 46.05) mm, rotated rx 94.06 ry 0 rz 180 deg; joints [-1.033, -84.136, 122.156, 178.324, 38.032, -174.624]
  MoveL 4940 to (0, -44.76, 46.05) mm, rotated rx 94.06 ry 0 rz 180 deg; joints [-0.882, -71.657, 106.698, 178.464, 35.051, -174.686]
  MoveL 4941 to (0, -44.79, 45.45) mm, rotated rx 91.73 ry 0 rz 180 deg; joints [-0.256, -71.738, 106.617, 179.552, 34.88, -177.898]
  MoveL 4942 to (-200, -44.79, 45.45) mm, rotated rx 91.73 ry 0 rz 180 deg; joints [-0.3, -84.232, 122.068, 179.511, 37.837, -177.88]
  MoveL 4943 to (-200, -44.8, 44.85) mm, rotated rx 90 ry 0 rz 180 deg; joints [0.257, -84.283, 122.01, -179.579, 37.728, 179.667]
  MoveL 4944 to (0, -44.8, 44.85) mm, rotated rx 90 ry 0 rz 180 deg; joints [0.22, -71.78, 106.562, -179.615, 34.783, 179.683]
  MoveL 4945 to (0, -44.8, 44.25) mm, rotated rx 90 ry 0 rz 180 deg; joints [0.245, -71.78, 106.562, -179.571, 34.783, 179.647]
  MoveL 4946 to (-200, -44.8, 44.25) mm, rotated rx 90 ry 0 rz 180 deg; joints [0.287, -84.282, 122.009, -179.531, 37.728, 179.629]
  MoveL 4947 to (-200, -44.8, 43.65) mm, rotated rx 90 ry 0 rz 180 deg; joints [0.316, -84.282, 122.009, -179.483, 37.728, 179.591]
  MoveL 4948 to (0, -44.8, 43.65) mm, rotated rx 90 ry 0 rz 180 deg; joints [0.27, -71.78, 106.562, -179.527, 34.783, 179.611]
  MoveL 4949 to (0, -44.8, 43.05) mm, rotated rx 90 ry 0 rz 180 deg; joints [0.295, -71.78, 106.562, -179.483, 34.783, 179.575]
  MoveL 4950 to (-200, -44.8, 43.05) mm, rotated rx 90 ry 0 rz 180 deg; joints [0.345, -84.282, 122.009, -179.436, 37.728, 179.554]
  MoveL 4951 to (-200, -44.8, 42.45) mm, rotated rx 90 ry 0 rz 180 deg; joints [0.375, -84.282, 122.009, -179.388, 37.729, 179.516]
  MoveL 4952 to (0, -44.8, 42.45) mm, rotated rx 90 ry 0 rz 180 deg; joints [0.32, -71.779, 106.561, -179.439, 34.783, 179.539]
  MoveL 4953 to (0, -44.8, 41.85) mm, rotated rx 90 ry 0 rz 180 deg; joints [0.345, -71.779, 106.561, -179.395, 34.783, 179.503]
  MoveL 4954 to (-200, -44.8, 41.85) mm, rotated rx 90 ry 0 rz 180 deg; joints [0.404, -84.281, 122.008, -179.34, 37.729, 179.478]
  MoveL 4955 to (-200, -44.8, 41.25) mm, rotated rx 90 ry 0 rz 180 deg; joints [0.433, -84.281, 122.008, -179.292, 37.729, 179.44]
  MoveL 4956 to (0, -44.8, 41.25) mm, rotated rx 90 ry 0 rz 180 deg; joints [0.37, -71.779, 106.561, -179.351, 34.784, 179.467]
  MoveL 4957 to (0, -44.8, 40.65) mm, rotated rx 90 ry 0 rz 180 deg; joints [0.395, -71.779, 106.56, -179.307, 34.784, 179.431]
  MoveL 4958 to (-200, -44.8, 40.65) mm, rotated rx 90 ry 0 rz 180 deg; joints [0.463, -84.281, 122.008, -179.244, 37.729, 179.402]
  MoveL 4959 to (-200, -44.8, 40.05) mm, rotated rx 90 ry 0 rz 180 deg; joints [0.492, -84.281, 122.007, -179.196, 37.73, 179.364]
  MoveL 4960 to (0, -44.8, 40.05) mm, rotated rx 90 ry 0 rz 180 deg; joints [0.42, -71.778, 106.56, -179.263, 34.784, 179.395]
  MoveL 4961 to (0, -44.8, 39.45) mm, rotated rx 90 ry 0 rz 180 deg; joints [0.445, -71.778, 106.56, -179.219, 34.784, 179.359]
  MoveL 4962 to (-200, -44.8, 39.45) mm, rotated rx 90 ry 0 rz 180 deg; joints [0.521, -84.28, 122.007, -179.148, 37.73, 179.326]
  MoveL 4963 to (-200, -44.8, 38.85) mm, rotated rx 90 ry 0 rz 180 deg; joints [0.551, -84.28, 122.007, -179.1, 37.73, 179.288]
  MoveL 4964 to (0, -44.8, 38.85) mm, rotated rx 90 ry 0 rz 180 deg; joints [0.47, -71.778, 106.559, -179.175, 34.784, 179.323]
  MoveL 4965 to (0, -44.8, 38.25) mm, rotated rx 90 ry 0 rz 180 deg; joints [0.495, -71.777, 106.559, -179.131, 34.784, 179.287]
  MoveL 4966 to (-200, -44.8, 38.25) mm, rotated rx 90 ry 0 rz 180 deg; joints [0.58, -84.279, 122.006, -179.052, 37.73, 179.25]
  MoveL 4967 to (-200, -44.8, 37.65) mm, rotated rx 90 ry 0 rz 180 deg; joints [0.609, -84.279, 122.006, -179.004, 37.731, 179.212]
  MoveL 4968 to (0, -44.8, 37.65) mm, rotated rx 90 ry 0 rz 180 deg; joints [0.521, -71.777, 106.558, -179.088, 34.785, 179.251]
  MoveL 4969 to (0, -44.8, 37.05) mm, rotated rx 90 ry 0 rz 180 deg; joints [0.546, -71.777, 106.558, -179.044, 34.785, 179.214]
  MoveL 4970 to (-200, -44.8, 37.05) mm, rotated rx 90 ry 0 rz 180 deg; joints [0.639, -84.279, 122.005, -178.956, 37.731, 179.174]
  MoveL 4971 to (-200, -44.8, 36.45) mm, rotated rx 90 ry 0 rz 180 deg; joints [0.668, -84.278, 122.005, -178.908, 37.732, 179.137]
  MoveL 4972 to (0, -44.8, 36.45) mm, rotated rx 90 ry 0 rz 180 deg; joints [0.571, -71.776, 106.557, -179, 34.785, 179.178]
  MoveL 4973 to (0, -44.8, 35.85) mm, rotated rx 90 ry 0 rz 180 deg; joints [0.596, -71.776, 106.557, -178.956, 34.785, 179.142]
  MoveL 4974 to (-200, -44.8, 35.85) mm, rotated rx 90 ry 0 rz 180 deg; joints [0.697, -84.278, 122.004, -178.86, 37.732, 179.099]
  MoveL 4975 to (-200, -44.8, 35.25) mm, rotated rx 90 ry 0 rz 180 deg; joints [0.727, -84.277, 122.004, -178.812, 37.732, 179.061]
  MoveL 4976 to (0, -44.8, 35.25) mm, rotated rx 90 ry 0 rz 180 deg; joints [0.621, -71.776, 106.556, -178.912, 34.786, 179.106]
  MoveL 4977 to (0, -44.8, 34.65) mm, rotated rx 90 ry 0 rz 180 deg; joints [0.646, -71.775, 106.556, -178.868, 34.786, 179.07]
  MoveL 4978 to (-200, -44.8, 34.65) mm, rotated rx 90 ry 0 rz 180 deg; joints [0.756, -84.277, 122.003, -178.765, 37.733, 179.023]
  MoveL 4979 to (-200, -44.8, 34.05) mm, rotated rx 90 ry 0 rz 180 deg; joints [0.785, -84.276, 122.003, -178.717, 37.733, 178.985]
  MoveL 4980 to (0, -44.8, 34.05) mm, rotated rx 90 ry 0 rz 180 deg; joints [0.671, -71.775, 106.555, -178.824, 34.786, 179.034]
  MoveL 4981 to (0, -44.8, 33.45) mm, rotated rx 90 ry 0 rz 180 deg; joints [0.696, -71.774, 106.555, -178.78, 34.786, 178.998]
  MoveL 4982 to (-200, -44.8, 33.45) mm, rotated rx 90 ry 0 rz 180 deg; joints [0.815, -84.276, 122.002, -178.669, 37.734, 178.947]
  MoveL 4983 to (-200, -44.8, 32.85) mm, rotated rx 90 ry 0 rz 180 deg; joints [0.844, -84.275, 122.001, -178.621, 37.734, 178.909]
  MoveL 4984 to (0, -44.8, 32.85) mm, rotated rx 90 ry 0 rz 180 deg; joints [0.721, -71.774, 106.554, -178.736, 34.787, 178.962]
  MoveL 4985 to (0, -44.8, 32.25) mm, rotated rx 90 ry 0 rz 180 deg; joints [0.746, -71.773, 106.553, -178.692, 34.787, 178.926]
  MoveL 4986 to (-200, -44.8, 32.25) mm, rotated rx 90 ry 0 rz 180 deg; joints [0.873, -84.275, 122.001, -178.573, 37.735, 178.871]
  MoveL 4987 to (-200, -44.8, 31.65) mm, rotated rx 90 ry 0 rz 180 deg; joints [0.903, -84.274, 122, -178.525, 37.735, 178.833]
  MoveL 4988 to (0, -44.8, 31.65) mm, rotated rx 90 ry 0 rz 180 deg; joints [0.771, -71.773, 106.553, -178.648, 34.787, 178.89]
  MoveL 4989 to (0, -44.8, 31.05) mm, rotated rx 90 ry 0 rz 180 deg; joints [0.796, -71.772, 106.552, -178.604, 34.788, 178.854]
  MoveL 4990 to (-200, -44.8, 31.05) mm, rotated rx 90 ry 0 rz 180 deg; joints [0.932, -84.273, 121.999, -178.477, 37.736, 178.796]
  MoveL 4991 to (-200, -44.8, 30.45) mm, rotated rx 90 ry 0 rz 180 deg; joints [0.961, -84.273, 121.999, -178.429, 37.736, 178.758]
  MoveL 4992 to (0, -44.8, 30.45) mm, rotated rx 90 ry 0 rz 180 deg; joints [0.821, -71.772, 106.551, -178.561, 34.788, 178.818]
  MoveL 4993 to (0, -44.8, 29.85) mm, rotated rx 90 ry 0 rz 180 deg; joints [0.846, -71.771, 106.551, -178.517, 34.788, 178.782]
  MoveL 4994 to (-200, -44.8, 29.85) mm, rotated rx 90 ry 0 rz 180 deg; joints [0.991, -84.272, 121.998, -178.381, 37.737, 178.72]
  MoveL 4995 to (-200, -44.8, 29.25) mm, rotated rx 90 ry 0 rz 180 deg; joints [1.02, -84.271, 121.997, -178.333, 37.737, 178.682]
  MoveL 4996 to (0, -44.8, 29.25) mm, rotated rx 90 ry 0 rz 180 deg; joints [0.871, -71.771, 106.55, -178.473, 34.789, 178.746]
  MoveL 4997 to (0, -44.8, 28.65) mm, rotated rx 90 ry 0 rz 180 deg; joints [0.896, -71.77, 106.549, -178.429, 34.789, 178.71]
  MoveL 4998 to (-200, -44.8, 28.65) mm, rotated rx 90 ry 0 rz 180 deg; joints [1.049, -84.271, 121.996, -178.285, 37.738, 178.644]
  MoveL 4999 to (-200, -44.8, 28.05) mm, rotated rx 90 ry 0 rz 180 deg; joints [1.079, -84.27, 121.996, -178.238, 37.739, 178.606]
  MoveL 5000 to (0, -44.8, 28.05) mm, rotated rx 90 ry 0 rz 180 deg; joints [0.921, -71.77, 106.548, -178.385, 34.789, 178.674]
  MoveL 5001 to (0, -44.8, 27.45) mm, rotated rx 90 ry 0 rz 180 deg; joints [0.946, -71.769, 106.548, -178.341, 34.79, 178.637]
  MoveL 5002 to (-200, -44.8, 27.45) mm, rotated rx 90 ry 0 rz 180 deg; joints [1.108, -84.269, 121.995, -178.19, 37.739, 178.568]
  MoveL 5003 to (-200, -44.8, 26.85) mm, rotated rx 90 ry 0 rz 180 deg; joints [1.137, -84.268, 121.994, -178.142, 37.74, 178.53]
  MoveL 5004 to (0, -44.8, 26.85) mm, rotated rx 90 ry 0 rz 180 deg; joints [0.971, -71.768, 106.547, -178.297, 34.79, 178.601]
  MoveL 5005 to (0, -44.8, 26.25) mm, rotated rx 90 ry 0 rz 180 deg; joints [0.997, -71.768, 106.546, -178.253, 34.79, 178.565]
  MoveL 5006 to (-200, -44.8, 26.25) mm, rotated rx 90 ry 0 rz 180 deg; joints [1.167, -84.268, 121.993, -178.094, 37.741, 178.492]
  MoveL 5007 to (-200, -44.8, 25.65) mm, rotated rx 90 ry 0 rz 180 deg; joints [1.196, -84.267, 121.992, -178.046, 37.741, 178.455]
  MoveL 5008 to (0, -44.8, 25.65) mm, rotated rx 90 ry 0 rz 180 deg; joints [1.022, -71.767, 106.545, -178.209, 34.791, 178.529]
  MoveL 5009 to (0, -44.8, 25.05) mm, rotated rx 90 ry 0 rz 180 deg; joints [1.047, -71.767, 106.544, -178.165, 34.791, 178.493]
  MoveL 5010 to (-200, -44.8, 25.05) mm, rotated rx 90 ry 0 rz 180 deg; joints [1.225, -84.266, 121.991, -177.998, 37.742, 178.417]
  MoveL 5011 to (-200, -44.8, 24.45) mm, rotated rx 90 ry 0 rz 180 deg; joints [1.255, -84.265, 121.99, -177.95, 37.743, 178.379]
  MoveL 5012 to (0, -44.8, 24.45) mm, rotated rx 90 ry 0 rz 180 deg; joints [1.072, -71.766, 106.543, -178.122, 34.792, 178.457]
  MoveL 5013 to (0, -44.8, 23.85) mm, rotated rx 90 ry 0 rz 180 deg; joints [1.097, -71.765, 106.542, -178.078, 34.792, 178.421]
  MoveL 5014 to (-200, -44.8, 23.85) mm, rotated rx 90 ry 0 rz 180 deg; joints [1.284, -84.264, 121.989, -177.902, 37.744, 178.341]
  MoveL 5015 to (-200, -44.8, 23.25) mm, rotated rx 90 ry 0 rz 180 deg; joints [1.313, -84.263, 121.988, -177.854, 37.744, 178.303]
  MoveL 5016 to (0, -44.8, 23.25) mm, rotated rx 90 ry 0 rz 180 deg; joints [1.122, -71.764, 106.541, -178.034, 34.793, 178.385]
  MoveL 5017 to (0, -44.8, 22.65) mm, rotated rx 90 ry 0 rz 180 deg; joints [1.147, -71.764, 106.54, -177.99, 34.793, 178.349]
  MoveL 5018 to (-200, -44.8, 22.65) mm, rotated rx 90 ry 0 rz 180 deg; joints [1.342, -84.263, 121.987, -177.807, 37.745, 178.265]
  MoveL 5019 to (-200, -44.8, 22.05) mm, rotated rx 90 ry 0 rz 180 deg; joints [1.372, -84.262, 121.986, -177.759, 37.746, 178.227]
  MoveL 5020 to (0, -44.8, 22.05) mm, rotated rx 90 ry 0 rz 180 deg; joints [1.172, -71.763, 106.539, -177.946, 34.794, 178.313]
  MoveL 5021 to (0, -44.8, 21.45) mm, rotated rx 90 ry 0 rz 180 deg; joints [1.197, -71.762, 106.538, -177.902, 34.794, 178.277]
  MoveL 5022 to (-200, -44.8, 21.45) mm, rotated rx 90 ry 0 rz 180 deg; joints [1.401, -84.261, 121.985, -177.711, 37.747, 178.19]
  MoveL 5023 to (-200, -44.8, 20.85) mm, rotated rx 90 ry 0 rz 180 deg; joints [1.43, -84.26, 121.984, -177.663, 37.747, 178.152]
  MoveL 5024 to (0, -44.8, 20.85) mm, rotated rx 90 ry 0 rz 180 deg; joints [1.222, -71.761, 106.537, -177.858, 34.794, 178.241]
  MoveL 5025 to (0, -44.8, 20.25) mm, rotated rx 90 ry 0 rz 180 deg; joints [1.247, -71.761, 106.536, -177.814, 34.795, 178.205]
  MoveL 5026 to (-200, -44.8, 20.25) mm, rotated rx 90 ry 0 rz 180 deg; joints [1.46, -84.259, 121.983, -177.615, 37.748, 178.114]
  MoveL 5027 to (-200, -44.8, 19.65) mm, rotated rx 90 ry 0 rz 180 deg; joints [1.489, -84.258, 121.982, -177.567, 37.749, 178.076]
  MoveL 5028 to (0, -44.8, 19.65) mm, rotated rx 90 ry 0 rz 180 deg; joints [1.272, -71.76, 106.535, -177.77, 34.795, 178.169]
  MoveL 5029 to (0, -44.8, 19.05) mm, rotated rx 90 ry 0 rz 180 deg; joints [1.297, -71.759, 106.534, -177.727, 34.796, 178.133]
  MoveL 5030 to (-200, -44.8, 19.05) mm, rotated rx 90 ry 0 rz 180 deg; joints [1.518, -84.257, 121.981, -177.519, 37.75, 178.038]
  MoveL 5031 to (-200, -44.8, 18.45) mm, rotated rx 90 ry 0 rz 180 deg; joints [1.548, -84.256, 121.98, -177.472, 37.751, 178]
  MoveL 5032 to (0, -44.8, 18.45) mm, rotated rx 90 ry 0 rz 180 deg; joints [1.322, -71.758, 106.533, -177.683, 34.797, 178.097]
  MoveL 5033 to (0, -44.8, 17.85) mm, rotated rx 90 ry 0 rz 180 deg; joints [1.347, -71.757, 106.532, -177.639, 34.797, 178.061]
  MoveL 5034 to (-200, -44.8, 17.85) mm, rotated rx 90 ry 0 rz 180 deg; joints [1.577, -84.255, 121.979, -177.424, 37.752, 177.962]
  MoveL 5035 to (-200, -44.8, 17.25) mm, rotated rx 90 ry 0 rz 180 deg; joints [1.606, -84.254, 121.977, -177.376, 37.753, 177.925]
  MoveL 5036 to (0, -44.8, 17.25) mm, rotated rx 90 ry 0 rz 180 deg; joints [1.372, -71.756, 106.53, -177.595, 34.798, 178.025]
  MoveL 5037 to (0, -44.8, 16.65) mm, rotated rx 90 ry 0 rz 180 deg; joints [1.397, -71.755, 106.529, -177.551, 34.798, 177.989]
  MoveL 5038 to (-200, -44.8, 16.65) mm, rotated rx 90 ry 0 rz 180 deg; joints [1.636, -84.253, 121.976, -177.328, 37.754, 177.887]
  MoveL 5039 to (-200, -44.8, 16.05) mm, rotated rx 90 ry 0 rz 180 deg; joints [1.665, -84.251, 121.975, -177.28, 37.755, 177.849]
  MoveL 5040 to (0, -44.8, 16.05) mm, rotated rx 90 ry 0 rz 180 deg; joints [1.422, -71.755, 106.528, -177.507, 34.799, 177.953]
  MoveL 5041 to (0, -44.8, 15.45) mm, rotated rx 90 ry 0 rz 180 deg; joints [1.447, -71.754, 106.527, -177.463, 34.799, 177.917]
  MoveL 5042 to (-200, -44.8, 15.45) mm, rotated rx 90 ry 0 rz 180 deg; joints [1.694, -84.25, 121.974, -177.232, 37.756, 177.811]
  MoveL 5043 to (-200, -44.8, 14.85) mm, rotated rx 89.41 ry 0 rz 180 deg; joints [1.903, -84.256, 121.947, -176.889, 37.732, 176.95]
  MoveL 5044 to (0, -44.8, 14.85) mm, rotated rx 89.41 ry 0 rz 180 deg; joints [1.626, -71.759, 106.501, -177.149, 34.776, 177.068]
  MoveL 5045 to (0, -44.78, 14.25) mm, rotated rx 87.09 ry 0 rz 180 deg; joints [2.258, -71.764, 106.41, -176.033, 34.711, 173.825]
  MoveL 5046 to (-200, -44.78, 14.25) mm, rotated rx 87.09 ry 0 rz 180 deg; joints [2.643, -84.261, 121.852, -175.673, 37.67, 173.661]
  MoveL 5047 to (-200, -44.74, 13.65) mm, rotated rx 84.77 ry 0 rz 180 deg; joints [3.383, -84.232, 121.768, -174.458, 37.665, 170.373]
  MoveL 5048 to (0, -44.74, 13.65) mm, rotated rx 84.77 ry 0 rz 180 deg; joints [2.891, -71.74, 106.328, -174.917, 34.693, 170.582]
  MoveL 5049 to (0, -44.67, 13.05) mm, rotated rx 82.44 ry 0 rz 180 deg; joints [3.524, -71.69, 106.255, -173.806, 34.722, 167.344]
  MoveL 5050 to (-200, -44.67, 13.05) mm, rotated rx 82.44 ry 0 rz 180 deg; joints [4.123, -84.17, 121.694, -173.251, 37.717, 167.094]
  MoveL 5051 to (-200, -44.58, 12.46) mm, rotated rx 80.12 ry 0 rz 180 deg; joints [4.861, -84.075, 121.631, -172.058, 37.823, 163.831]
  MoveL 5052 to (0, -44.58, 12.46) mm, rotated rx 80.12 ry 0 rz 180 deg; joints [4.155, -71.611, 106.191, -172.706, 34.798, 164.12]
  MoveL 5053 to (0, -44.47, 11.87) mm, rotated rx 77.8 ry 0 rz 180 deg; joints [4.784, -71.505, 106.136, -171.622, 34.919, 160.912]
  MoveL 5054 to (-200, -44.47, 11.87) mm, rotated rx 77.8 ry 0 rz 180 deg; joints [5.595, -83.947, 121.578, -170.884, 37.984, 160.589]
  MoveL 5055 to (-200, -44.33, 11.29) mm, rotated rx 75.47 ry 0 rz 180 deg; joints [6.326, -83.786, 121.537, -169.737, 38.199, 157.376]
  MoveL 5056 to (0, -44.33, 11.29) mm, rotated rx 75.47 ry 0 rz 180 deg; joints [5.409, -71.372, 106.091, -170.56, 35.085, 157.726]
  MoveL 5057 to (0, -44.16, 10.71) mm, rotated rx 73.15 ry 0 rz 180 deg; joints [6.03, -71.212, 106.054, -169.525, 35.295, 154.569]
  MoveL 5058 to (-200, -44.16, 10.71) mm, rotated rx 73.15 ry 0 rz 180 deg; joints [7.049, -83.593, 121.505, -168.621, 38.465, 154.196]
  MoveL 5059 to (-200, -43.98, 10.14) mm, rotated rx 70.83 ry 0 rz 180 deg; joints [7.766, -83.368, 121.485, -167.542, 38.782, 151.056]
  MoveL 5060 to (0, -43.98, 10.14) mm, rotated rx 70.83 ry 0 rz 180 deg; joints [6.645, -71.025, 106.027, -168.52, 35.548, 151.445]
  MoveL 5061 to (0, -43.77, 9.58) mm, rotated rx 68.51 ry 0 rz 180 deg; joints [7.252, -70.812, 106.009, -167.55, 35.842, 148.359]
  MoveL 5062 to (-200, -43.77, 9.58) mm, rotated rx 68.51 ry 0 rz 180 deg; joints [8.473, -83.112, 121.475, -166.503, 39.147, 147.961]
  MoveL 5063 to (-200, -43.54, 9.02) mm, rotated rx 66.18 ry 0 rz 180 deg; joints [9.171, -82.824, 121.475, -165.508, 39.558, 144.913]
  MoveL 5064 to (0, -43.54, 9.02) mm, rotated rx 66.18 ry 0 rz 180 deg; joints [7.852, -70.573, 106, -166.618, 36.176, 145.312]
  MoveL 5065 to (0, -43.29, 8.48) mm, rotated rx 63.86 ry 0 rz 180 deg; joints [8.442, -70.308, 106, -165.727, 36.548, 142.31]
  MoveL 5066 to (-200, -43.29, 8.48) mm, rotated rx 63.86 ry 0 rz 180 deg; joints [9.857, -82.506, 121.485, -164.559, 40.013, 141.915]
  MoveL 5067 to (-200, -43.01, 7.95) mm, rotated rx 61.54 ry 0 rz 180 deg; joints [10.53, -82.157, 121.505, -163.66, 40.511, 138.971]
  MoveL 5068 to (0, -43.01, 7.95) mm, rotated rx 61.54 ry 0 rz 180 deg; joints [9.022, -70.018, 106.009, -164.88, 36.956, 139.353]
  MoveL 5069 to (0, -42.71, 7.42) mm, rotated rx 59.21 ry 0 rz 180 deg; joints [9.591, -69.703, 106.026, -164.077, 37.399, 136.444]
  MoveL 5070 to (-200, -42.71, 7.42) mm, rotated rx 59.21 ry 0 rz 180 deg; joints [11.19, -81.779, 121.535, -162.812, 41.048, 136.083]
  MoveL 5071 to (-200, -42.4, 6.92) mm, rotated rx 56.89 ry 0 rz 180 deg; joints [11.835, -81.372, 121.574, -162.015, 41.622, 133.252]
  MoveL 5072 to (0, -42.4, 6.92) mm, rotated rx 56.89 ry 0 rz 180 deg; joints [10.148, -69.364, 106.051, -163.322, 37.874, 133.587]
  MoveL 5073 to (0, -42.06, 6.42) mm, rotated rx 54.57 ry 0 rz 180 deg; joints [10.692, -69, 106.084, -162.613, 38.381, 130.778]
  MoveL 5074 to (-200, -42.06, 6.42) mm, rotated rx 54.57 ry 0 rz 180 deg; joints [12.464, -80.935, 121.621, -161.271, 42.232, 130.477]
  MoveL 5075 to (-200, -41.7, 5.94) mm, rotated rx 52.25 ry 0 rz 180 deg; joints [13.076, -80.471, 121.677, -160.578, 42.875, 127.758]
  MoveL 5076 to (0, -41.7, 5.94) mm, rotated rx 52.25 ry 0 rz 180 deg; joints [11.222, -68.614, 106.125, -161.952, 38.916, 128.02]
  MoveL 5077 to (0, -41.33, 5.47) mm, rotated rx 49.92 ry 0 rz 180 deg; joints [11.737, -68.204, 106.173, -161.339, 39.478, 125.313]
  MoveL 5078 to (-200, -41.33, 5.47) mm, rotated rx 49.92 ry 0 rz 180 deg; joints [13.671, -79.98, 121.741, -159.938, 43.548, 125.097]
  MoveL 5079 to (-200, -40.93, 5.02) mm, rotated rx 47.6 ry 0 rz 180 deg; joints [14.247, -79.462, 121.812, -159.349, 44.249, 122.492]
  MoveL 5080 to (0, -40.93, 5.02) mm, rotated rx 47.6 ry 0 rz 180 deg; joints [12.237, -67.772, 106.228, -160.774, 40.066, 122.656]
  MoveL 5081 to (0, -40.52, 4.59) mm, rotated rx 45.28 ry 0 rz 180 deg; joints [12.721, -67.319, 106.289, -160.255, 40.678, 120.049]
  MoveL 5082 to (-200, -40.52, 4.59) mm, rotated rx 45.28 ry 0 rz 180 deg; joints [14.803, -78.918, 121.891, -158.809, 44.977, 119.941]
  MoveL 5083 to (-200, -40.09, 4.17) mm, rotated rx 42.95 ry 0 rz 180 deg; joints [15.339, -78.349, 121.977, -158.319, 45.729, 117.445]
  MoveL 5084 to (0, -40.09, 4.17) mm, rotated rx 42.95 ry 0 rz 180 deg; joints [13.188, -66.844, 106.357, -159.782, 41.311, 117.492]
  MoveL 5085 to (0, -39.64, 3.77) mm, rotated rx 40.63 ry 0 rz 180 deg; joints [13.637, -66.349, 106.43, -159.354, 41.964, 114.981]
  MoveL 5086 to (-200, -39.64, 3.77) mm, rotated rx 40.63 ry 0 rz 180 deg; joints [15.855, -77.755, 122.068, -157.876, 46.504, 114.999]
  MoveL 5087 to (-200, -39.17, 3.39) mm, rotated rx 38.31 ry 0 rz 180 deg; joints [16.349, -77.137, 122.166, -157.478, 47.299, 112.602]
  MoveL 5088 to (0, -39.17, 3.39) mm, rotated rx 38.31 ry 0 rz 180 deg; joints [14.068, -65.834, 106.509, -158.969, 42.636, 112.515]
  MoveL 5089 to (0, -38.7, 3.02) mm, rotated rx 35.99 ry 0 rz 180 deg; joints [14.48, -65.3, 106.593, -158.627, 43.325, 110.094]
  MoveL 5090 to (-200, -38.7, 3.02) mm, rotated rx 35.99 ry 0 rz 180 deg; joints [16.821, -76.496, 122.268, -157.125, 48.112, 110.254]
  MoveL 5091 to (-200, -38.2, 2.68) mm, rotated rx 33.66 ry 0 rz 180 deg; joints [17.271, -75.833, 122.376, -156.814, 48.943, 107.95]
  MoveL 5092 to (0, -38.2, 2.68) mm, rotated rx 33.66 ry 0 rz 180 deg; joints [14.874, -64.748, 106.682, -158.326, 44.029, 107.716]
  MoveL 5093 to (0, -37.7, 2.36) mm, rotated rx 31.34 ry 0 rz 180 deg; joints [15.247, -64.178, 106.774, -158.064, 44.746, 105.379]
  MoveL 5094 to (-200, -37.7, 2.36) mm, rotated rx 31.34 ry 0 rz 180 deg; joints [17.697, -75.149, 122.487, -156.543, 49.789, 105.691]
  MoveL 5095 to (-200, -37.18, 2.06) mm, rotated rx 29.02 ry 0 rz 180 deg; joints [18.1, -74.444, 122.602, -156.311, 50.649, 103.472]
  MoveL 5096 to (0, -37.18, 2.06) mm, rotated rx 29.02 ry 0 rz 180 deg; joints [15.6, -63.591, 106.871, -157.84, 45.477, 103.08]
  MoveL 5097 to (0, -36.65, 1.78) mm, rotated rx 26.7 ry 0 rz 180 deg; joints [15.933, -62.988, 106.971, -157.653, 46.219, 100.817]
  MoveL 5098 to (-200, -36.65, 1.78) mm, rotated rx 26.7 ry 0 rz 180 deg; joints [18.48, -73.72, 122.721, -156.116, 51.522, 101.291]
  MoveL 5099 to (-200, -36.11, 1.52) mm, rotated rx 24.37 ry 0 rz 180 deg; joints [18.835, -72.976, 122.842, -155.956, 52.406, 99.146]
  MoveL 5100 to (0, -36.11, 1.52) mm, rotated rx 24.37 ry 0 rz 180 deg; joints [16.245, -62.37, 107.074, -157.5, 46.971, 98.589]
  MoveL 5101 to (0, -35.56, 1.28) mm, rotated rx 22.05 ry 0 rz 180 deg; joints [16.536, -61.737, 107.179, -157.38, 47.731, 96.394]
  MoveL 5102 to (-200, -35.56, 1.28) mm, rotated rx 22.05 ry 0 rz 180 deg; joints [19.165, -72.215, 122.966, -155.829, 53.3, 97.035]
  MoveL 5103 to (-200, -34.99, 1.07) mm, rotated rx 19.73 ry 0 rz 180 deg; joints [19.471, -71.437, 123.091, -155.735, 54.202, 94.955]
  MoveL 5104 to (0, -34.99, 1.07) mm, rotated rx 19.73 ry 0 rz 180 deg; joints [16.805, -61.09, 107.287, -157.293, 48.499, 94.229]
  MoveL 5105 to (0, -34.43, 0.88) mm, rotated rx 17.4 ry 0 rz 180 deg; joints [17.052, -60.431, 107.396, -157.236, 49.274, 92.093]
  MoveL 5106 to (-200, -34.43, 0.88) mm, rotated rx 17.4 ry 0 rz 180 deg; joints [19.751, -70.643, 123.218, -155.67, 55.112, 92.904]
  MoveL 5107 to (-200, -33.85, 0.71) mm, rotated rx 15.08 ry 0 rz 180 deg; joints [20.007, -69.835, 123.345, -155.635, 56.028, 90.88]
  MoveL 5108 to (0, -33.85, 0.71) mm, rotated rx 15.08 ry 0 rz 180 deg; joints [17.277, -59.759, 107.507, -157.208, 50.054, 89.983]
  MoveL 5109 to (0, -33.27, 0.56) mm, rotated rx 12.76 ry 0 rz 180 deg; joints [17.48, -59.076, 107.618, -157.208, 50.839, 87.897]
  MoveL 5110 to (-200, -33.27, 0.56) mm, rotated rx 12.76 ry 0 rz 180 deg; joints [20.237, -69.012, 123.474, -155.627, 56.95, 88.88]
  MoveL 5111 to (-200, -32.68, 0.45) mm, rotated rx 10.44 ry 0 rz 180 deg; joints [20.441, -68.177, 123.602, -155.646, 57.876, 86.901]
  MoveL 5112 to (0, -32.68, 0.45) mm, rotated rx 10.44 ry 0 rz 180 deg; joints [17.66, -58.383, 107.73, -157.235, 51.627, 85.834]
  MoveL 5113 to (0, -32.09, 0.35) mm, rotated rx 8.11 ry 0 rz 180 deg; joints [17.818, -57.682, 107.843, -157.287, 52.418, 83.792]
  MoveL 5114 to (-200, -32.09, 0.35) mm, rotated rx 8.11 ry 0 rz 180 deg; joints [20.619, -67.33, 123.729, -155.69, 58.805, 84.944]
  MoveL 5115 to (-200, -31.49, 0.28) mm, rotated rx 5.79 ry 0 rz 180 deg; joints [20.772, -66.472, 123.856, -155.757, 59.737, 83.004]
  MoveL 5116 to (0, -31.49, 0.28) mm, rotated rx 5.79 ry 0 rz 180 deg; joints [17.953, -56.971, 107.956, -157.363, 53.21, 81.768]
  MoveL 5117 to (0, -30.89, 0.23) mm, rotated rx 3.47 ry 0 rz 180 deg; joints [18.065, -56.254, 108.068, -157.463, 54.003, 79.761]
  MoveL 5118 to (-200, -30.89, 0.23) mm, rotated rx 3.47 ry 0 rz 180 deg; joints [20.898, -65.605, 123.982, -155.848, 60.67, 81.079]
